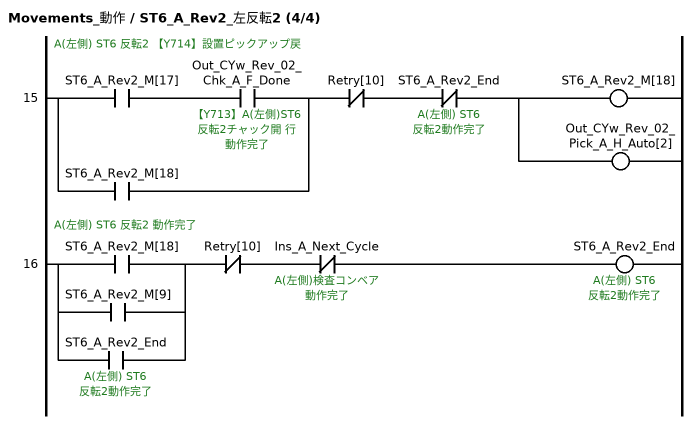
(* [picture p48: Movements_動作 / ST6_A_Rev2_左反転2, rungs 15-16] *)
(* Rung 15: A(左側) ST6 反転2 【Y714】設置ピックアップ戻 *)
_p89 := ((ST6_A_Rev2_M[17] AND Out_CYw_Rev_02_Chk_A_F_Done) OR ST6_A_Rev2_M[18]) AND NOT Retry[10] AND NOT ST6_A_Rev2_End;
ST6_A_Rev2_M[18] := _p89;
Out_CYw_Rev_02_Pick_A_H_Auto[2] := _p89;
(* Rung 16: A(左側) ST6 反転2 動作完了 *)
ST6_A_Rev2_End := (ST6_A_Rev2_M[18] OR ST6_A_Rev2_M[9] OR ST6_A_Rev2_End) AND NOT Retry[10] AND NOT Ins_A_Next_Cycle;

(* Section ST7_A_Dis2_左SF排出: ladder, written here as Structured Text *)

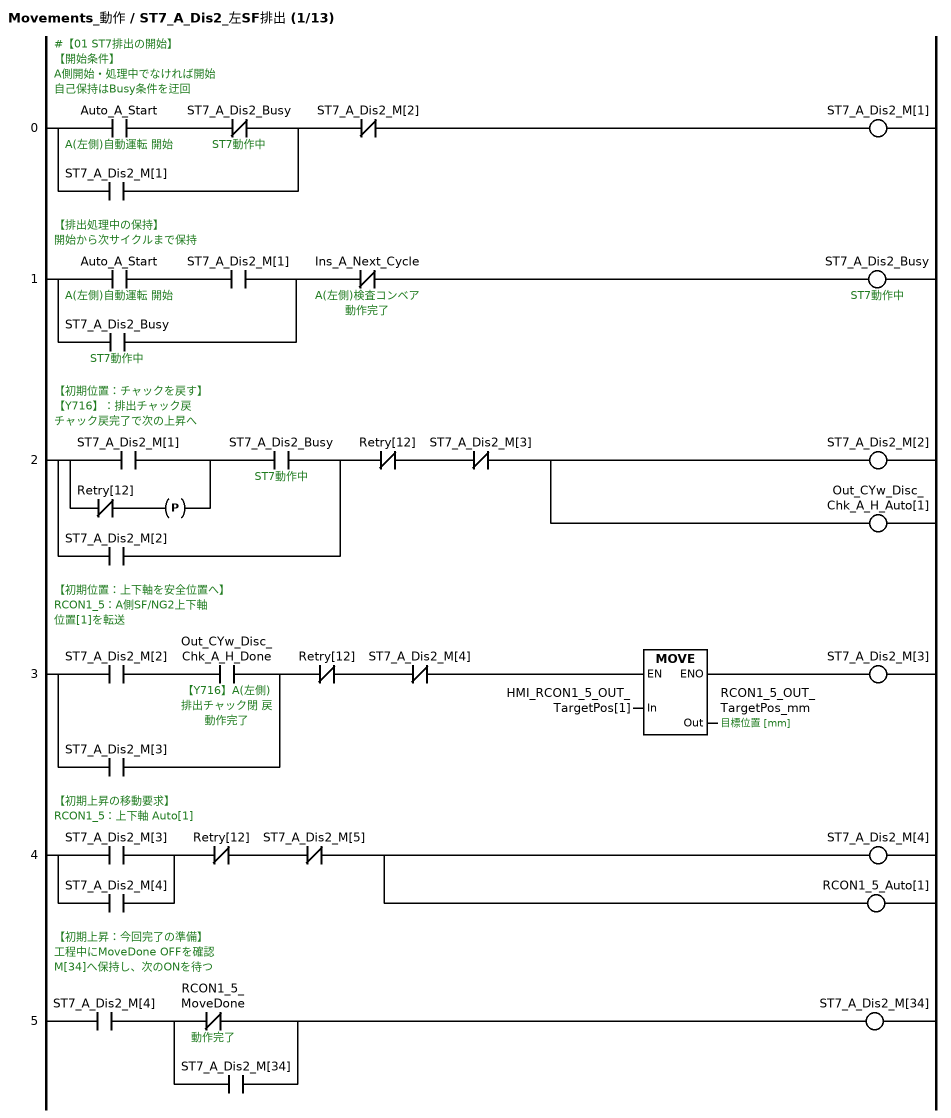
(* Rung 0: #【01 ST7排出の開始】 / 【開始条件】 / A側開始・処理中でなければ開始 / 自己保持はBusy条件を迂回 *)
ST7_A_Dis2_M[1] := ((Auto_A_Start AND NOT ST7_A_Dis2_Busy) OR ST7_A_Dis2_M[1]) AND NOT ST7_A_Dis2_M[2];
(* Rung 1: 【排出処理中の保持】 / 開始から次サイクルまで保持 *)
ST7_A_Dis2_Busy := ((Auto_A_Start AND ST7_A_Dis2_M[1]) OR ST7_A_Dis2_Busy) AND NOT Ins_A_Next_Cycle;
(* Rung 2: 【初期位置：チャックを戻す】 / 【Y716】：排出チャック戻 / チャック戻完了で次の上昇へ *)
_e90(CLK := NOT Retry[12]);
_p91 := (((ST7_A_Dis2_M[1] OR _e90.Q) AND ST7_A_Dis2_Busy) OR ST7_A_Dis2_M[2]) AND NOT Retry[12] AND NOT ST7_A_Dis2_M[3];
ST7_A_Dis2_M[2] := _p91;
Out_CYw_Disc_Chk_A_H_Auto[1] := _p91;
(* Rung 3: 【初期位置：上下軸を安全位置へ】 / RCON1_5：A側SF/NG2上下軸 / 位置[1]を転送 *)
IF ((ST7_A_Dis2_M[2] AND Out_CYw_Disc_Chk_A_H_Done) OR ST7_A_Dis2_M[3]) AND NOT Retry[12] AND NOT ST7_A_Dis2_M[4] THEN
    RCON1_5_OUT_TargetPos_mm := HMI_RCON1_5_OUT_TargetPos[1];
END_IF;
ST7_A_Dis2_M[3] := ((ST7_A_Dis2_M[2] AND Out_CYw_Disc_Chk_A_H_Done) OR ST7_A_Dis2_M[3]) AND NOT Retry[12] AND NOT ST7_A_Dis2_M[4];
(* Rung 4: 【初期上昇の移動要求】 / RCON1_5：上下軸 Auto[1] *)
_p92 := (ST7_A_Dis2_M[3] OR ST7_A_Dis2_M[4]) AND NOT Retry[12] AND NOT ST7_A_Dis2_M[5];
ST7_A_Dis2_M[4] := _p92;
RCON1_5_Auto[1] := _p92;
(* Rung 5: 【初期上昇：今回完了の準備】 / 工程中にMoveDone OFFを確認 / M[34]へ保持し、次のONを待つ *)
ST7_A_Dis2_M[34] := ST7_A_Dis2_M[4] AND (NOT RCON1_5_MoveDone OR ST7_A_Dis2_M[34]);

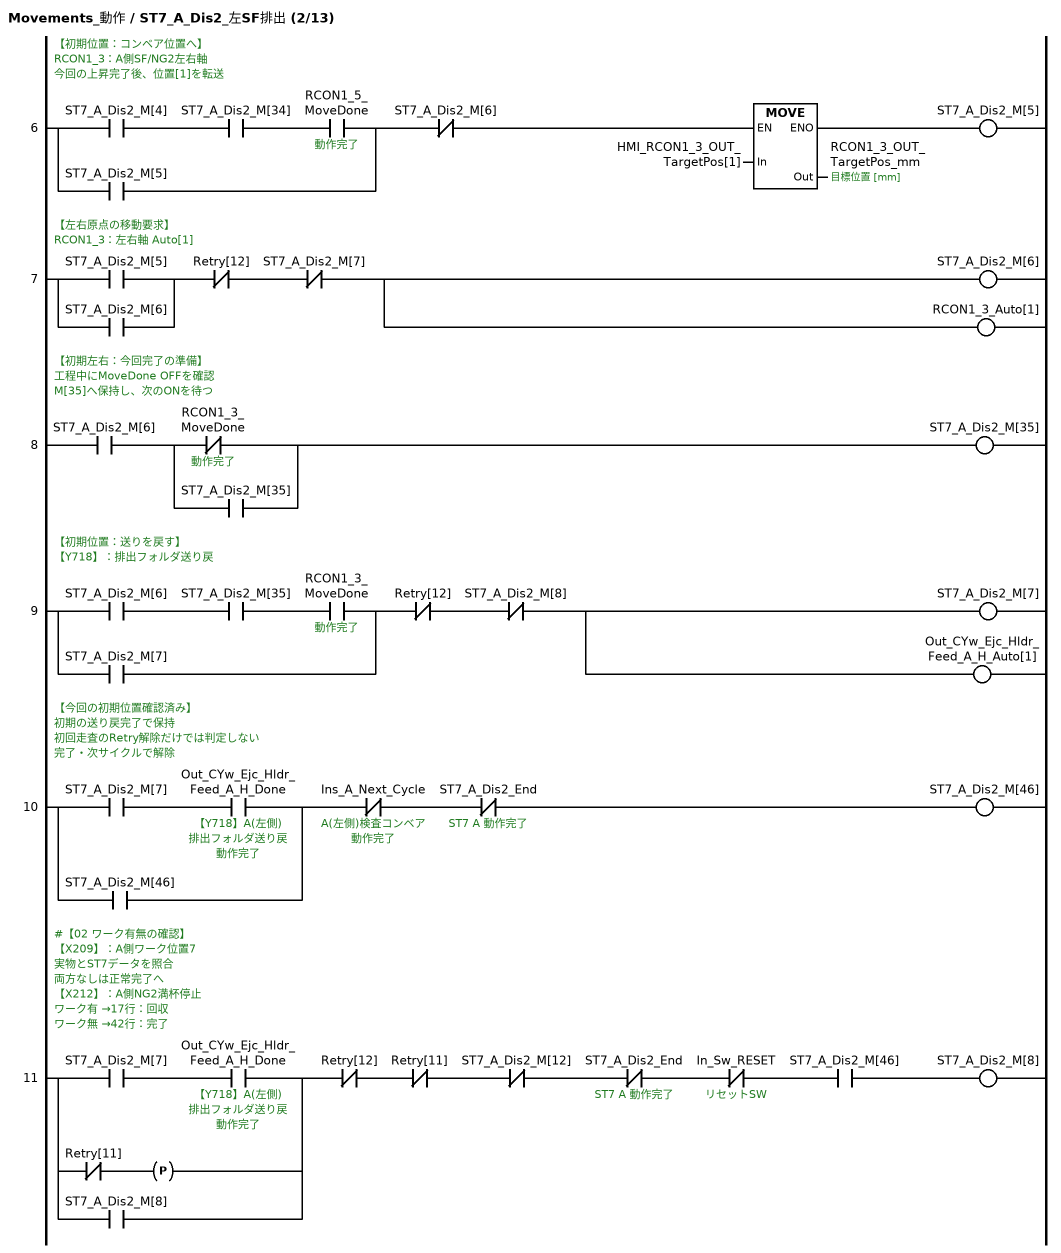
(* Rung 6: 【初期位置：コンベア位置へ】 / RCON1_3：A側SF/NG2左右軸 / 今回の上昇完了後、位置[1]を転送 *)
IF ((ST7_A_Dis2_M[4] AND ST7_A_Dis2_M[34] AND RCON1_5_MoveDone) OR ST7_A_Dis2_M[5]) AND NOT ST7_A_Dis2_M[6] THEN
    RCON1_3_OUT_TargetPos_mm := HMI_RCON1_3_OUT_TargetPos[1];
END_IF;
ST7_A_Dis2_M[5] := ((ST7_A_Dis2_M[4] AND ST7_A_Dis2_M[34] AND RCON1_5_MoveDone) OR ST7_A_Dis2_M[5]) AND NOT ST7_A_Dis2_M[6];
(* Rung 7: 【左右原点の移動要求】 / RCON1_3：左右軸 Auto[1] *)
_p93 := (ST7_A_Dis2_M[5] OR ST7_A_Dis2_M[6]) AND NOT Retry[12] AND NOT ST7_A_Dis2_M[7];
ST7_A_Dis2_M[6] := _p93;
RCON1_3_Auto[1] := _p93;
(* Rung 8: 【初期左右：今回完了の準備】 / 工程中にMoveDone OFFを確認 / M[35]へ保持し、次のONを待つ *)
ST7_A_Dis2_M[35] := ST7_A_Dis2_M[6] AND (NOT RCON1_3_MoveDone OR ST7_A_Dis2_M[35]);
(* Rung 9: 【初期位置：送りを戻す】 / 【Y718】：排出フォルダ送り戻 *)
_p94 := ((ST7_A_Dis2_M[6] AND ST7_A_Dis2_M[35] AND RCON1_3_MoveDone) OR ST7_A_Dis2_M[7]) AND NOT Retry[12] AND NOT ST7_A_Dis2_M[8];
ST7_A_Dis2_M[7] := _p94;
Out_CYw_Ejc_Hldr_Feed_A_H_Auto[1] := _p94;
(* Rung 10: 【今回の初期位置確認済み】 / 初期の送り戻完了で保持 / 初回走査のRetry解除だけでは判定しない / 完了・次サイクルで解除 *)
ST7_A_Dis2_M[46] := ((ST7_A_Dis2_M[7] AND Out_CYw_Ejc_Hldr_Feed_A_H_Done) OR ST7_A_Dis2_M[46]) AND NOT Ins_A_Next_Cycle AND NOT ST7_A_Dis2_End;
(* Rung 11: #【02 ワーク有無の確認】 / 【X209】：A側ワーク位置7 / 実物とST7データを照合 / 両方なしは正常完了へ / 【X212】：A側NG2満杯停止 / ワーク有 →17行：回収 / ワーク無 →42行：完了 *)
_e95(CLK := NOT Retry[11]);
ST7_A_Dis2_M[8] := ((ST7_A_Dis2_M[7] AND Out_CYw_Ejc_Hldr_Feed_A_H_Done) OR _e95.Q OR ST7_A_Dis2_M[8]) AND NOT Retry[12] AND NOT Retry[11] AND NOT ST7_A_Dis2_M[12] AND NOT ST7_A_Dis2_End AND NOT In_Sw_RESET AND ST7_A_Dis2_M[46];

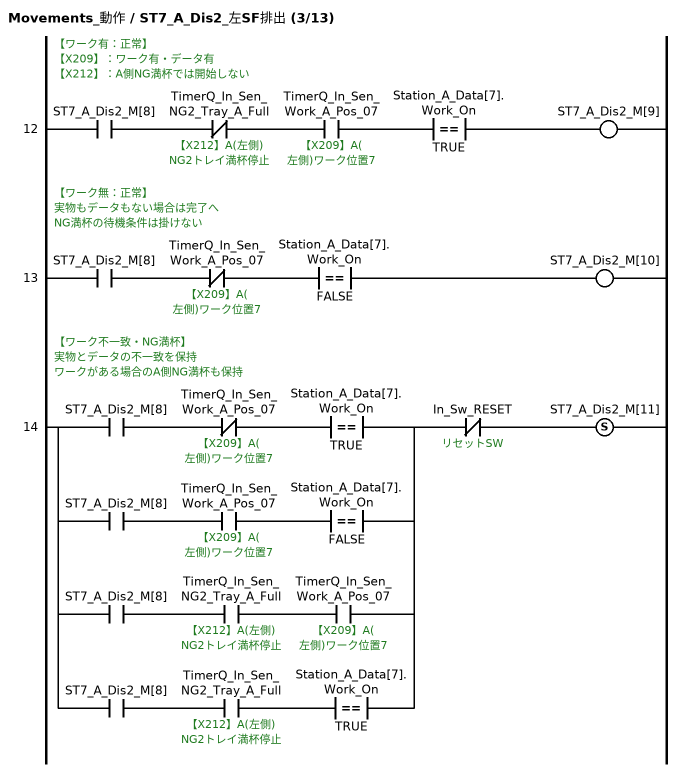
(* Rung 12: 【ワーク有：正常】 / 【X209】：ワーク有・データ有 / 【X212】：A側NG満杯では開始しない *)
ST7_A_Dis2_M[9] := ST7_A_Dis2_M[8] AND NOT TimerQ_In_Sen_NG2_Tray_A_Full AND TimerQ_In_Sen_Work_A_Pos_07 AND (Station_A_Data[7].Work_On = TRUE);
(* Rung 13: 【ワーク無：正常】 / 実物もデータもない場合は完了へ / NG満杯の待機条件は掛けない *)
ST7_A_Dis2_M[10] := ST7_A_Dis2_M[8] AND NOT TimerQ_In_Sen_Work_A_Pos_07 AND (Station_A_Data[7].Work_On = FALSE);
(* Rung 14: 【ワーク不一致・NG満杯】 / 実物とデータの不一致を保持 / ワークがある場合のA側NG満杯も保持 *)
IF ((ST7_A_Dis2_M[8] AND NOT TimerQ_In_Sen_Work_A_Pos_07 AND (Station_A_Data[7].Work_On = TRUE)) OR (ST7_A_Dis2_M[8] AND TimerQ_In_Sen_Work_A_Pos_07 AND (Station_A_Data[7].Work_On = FALSE)) OR (ST7_A_Dis2_M[8] AND TimerQ_In_Sen_NG2_Tray_A_Full AND TimerQ_In_Sen_Work_A_Pos_07) OR (ST7_A_Dis2_M[8] AND TimerQ_In_Sen_NG2_Tray_A_Full AND (Station_A_Data[7].Work_On = TRUE))) AND NOT In_Sw_RESET THEN
    ST7_A_Dis2_M[11] := TRUE;
END_IF;

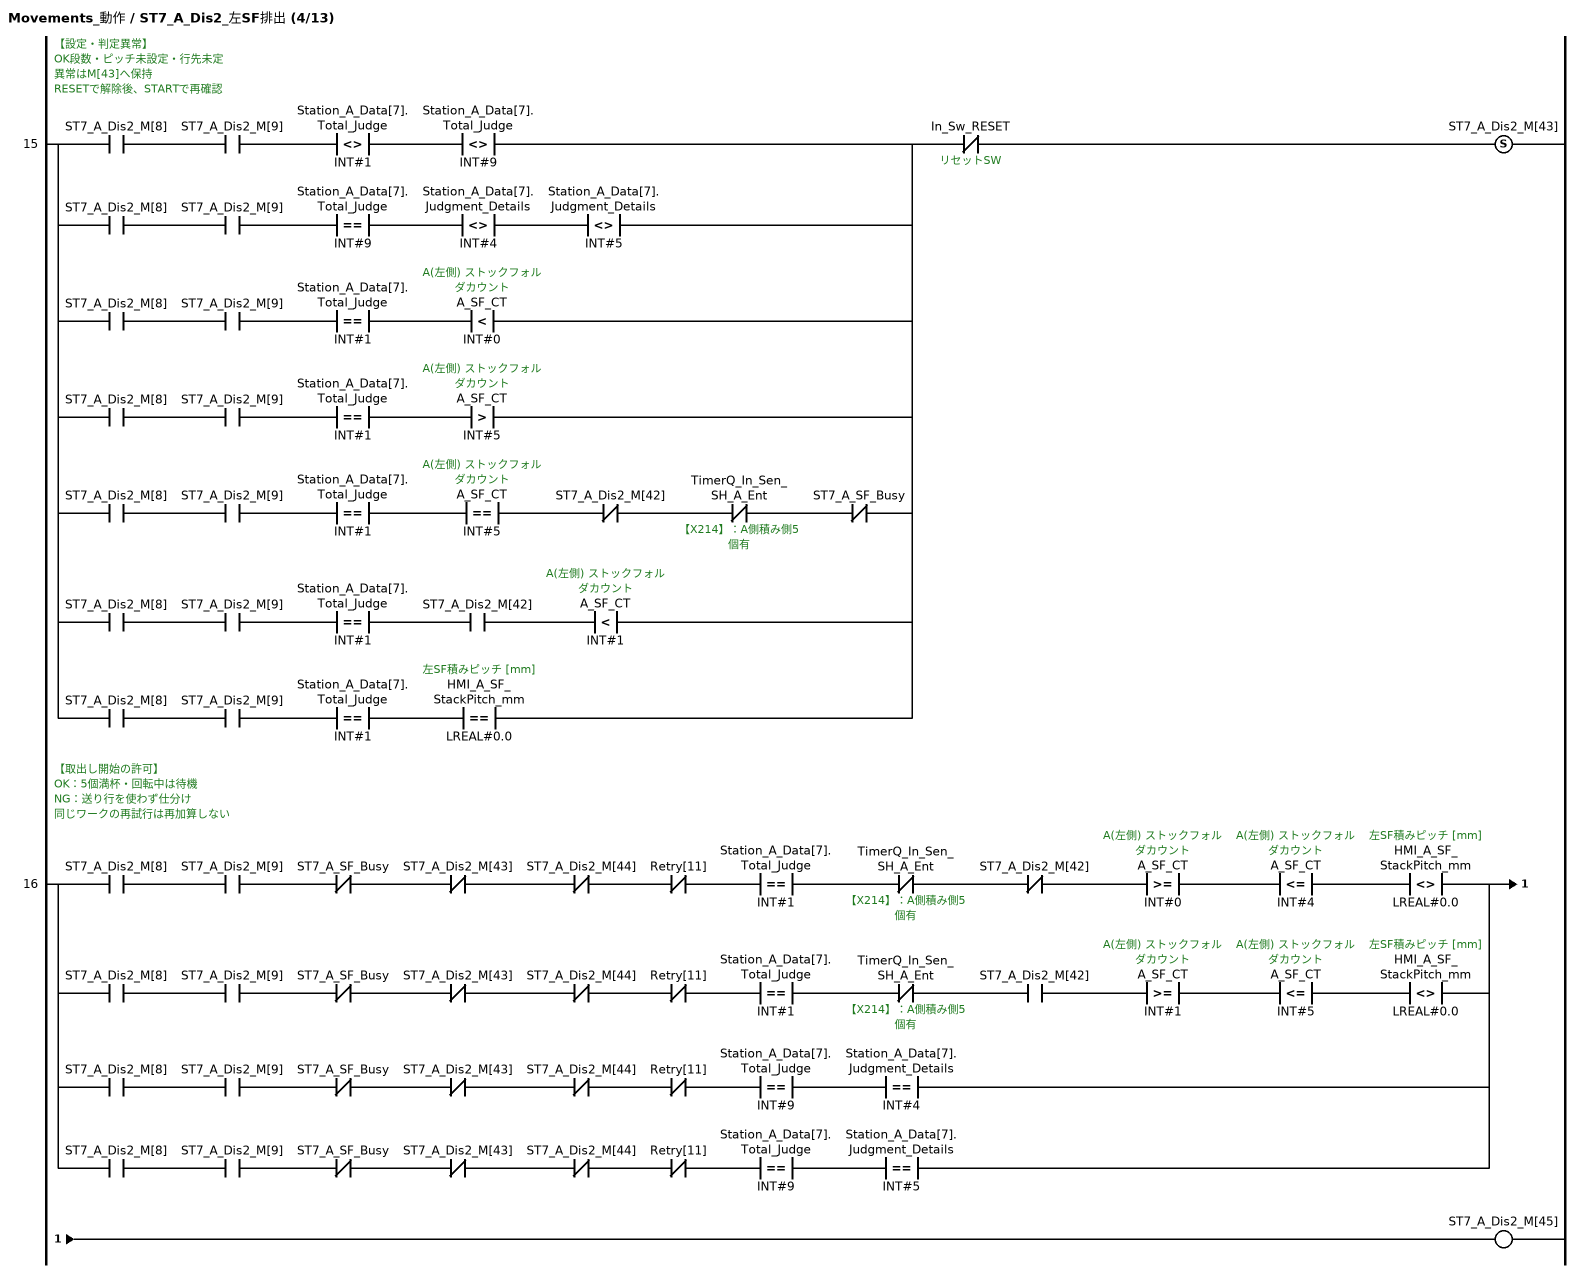
(* Rung 15: 【設定・判定異常】 / OK段数・ピッチ未設定・行先未定 / 異常はM[43]へ保持 / RESETで解除後、STARTで再確認 *)
IF ((ST7_A_Dis2_M[8] AND ST7_A_Dis2_M[9] AND (Station_A_Data[7].Total_Judge <> INT#1) AND (Station_A_Data[7].Total_Judge <> INT#9)) OR (ST7_A_Dis2_M[8] AND ST7_A_Dis2_M[9] AND (Station_A_Data[7].Total_Judge = INT#9) AND (Station_A_Data[7].Judgment_Details <> INT#4) AND (Station_A_Data[7].Judgment_Details <> INT#5)) OR (ST7_A_Dis2_M[8] AND ST7_A_Dis2_M[9] AND (Station_A_Data[7].Total_Judge = INT#1) AND (A_SF_CT < INT#0)) OR (ST7_A_Dis2_M[8] AND ST7_A_Dis2_M[9] AND (Station_A_Data[7].Total_Judge = INT#1) AND (A_SF_CT > INT#5)) OR (ST7_A_Dis2_M[8] AND ST7_A_Dis2_M[9] AND (Station_A_Data[7].Total_Judge = INT#1) AND (A_SF_CT = INT#5) AND NOT ST7_A_Dis2_M[42] AND NOT TimerQ_In_Sen_SH_A_Ent AND NOT ST7_A_SF_Busy) OR (ST7_A_Dis2_M[8] AND ST7_A_Dis2_M[9] AND (Station_A_Data[7].Total_Judge = INT#1) AND ST7_A_Dis2_M[42] AND (A_SF_CT < INT#1)) OR (ST7_A_Dis2_M[8] AND ST7_A_Dis2_M[9] AND (Station_A_Data[7].Total_Judge = INT#1) AND (HMI_A_SF_StackPitch_mm = LREAL#0.0))) AND NOT In_Sw_RESET THEN
    ST7_A_Dis2_M[43] := TRUE;
END_IF;
(* Rung 16: 【取出し開始の許可】 / OK：5個満杯・回転中は待機 / NG：送り行を使わず仕分け / 同じワークの再試行は再加算しない *)
ST7_A_Dis2_M[45] := (ST7_A_Dis2_M[8] AND ST7_A_Dis2_M[9] AND NOT ST7_A_SF_Busy AND NOT ST7_A_Dis2_M[43] AND NOT ST7_A_Dis2_M[44] AND NOT Retry[11] AND (Station_A_Data[7].Total_Judge = INT#1) AND NOT TimerQ_In_Sen_SH_A_Ent AND NOT ST7_A_Dis2_M[42] AND (A_SF_CT >= INT#0) AND (A_SF_CT <= INT#4) AND (HMI_A_SF_StackPitch_mm <> LREAL#0.0)) OR (ST7_A_Dis2_M[8] AND ST7_A_Dis2_M[9] AND NOT ST7_A_SF_Busy AND NOT ST7_A_Dis2_M[43] AND NOT ST7_A_Dis2_M[44] AND NOT Retry[11] AND (Station_A_Data[7].Total_Judge = INT#1) AND NOT TimerQ_In_Sen_SH_A_Ent AND ST7_A_Dis2_M[42] AND (A_SF_CT >= INT#1) AND (A_SF_CT <= INT#5) AND (HMI_A_SF_StackPitch_mm <> LREAL#0.0)) OR (ST7_A_Dis2_M[8] AND ST7_A_Dis2_M[9] AND NOT ST7_A_SF_Busy AND NOT ST7_A_Dis2_M[43] AND NOT ST7_A_Dis2_M[44] AND NOT Retry[11] AND (Station_A_Data[7].Total_Judge = INT#9) AND (Station_A_Data[7].Judgment_Details = INT#4)) OR (ST7_A_Dis2_M[8] AND ST7_A_Dis2_M[9] AND NOT ST7_A_SF_Busy AND NOT ST7_A_Dis2_M[43] AND NOT ST7_A_Dis2_M[44] AND NOT Retry[11] AND (Station_A_Data[7].Total_Judge = INT#9) AND (Station_A_Data[7].Judgment_Details = INT#5));

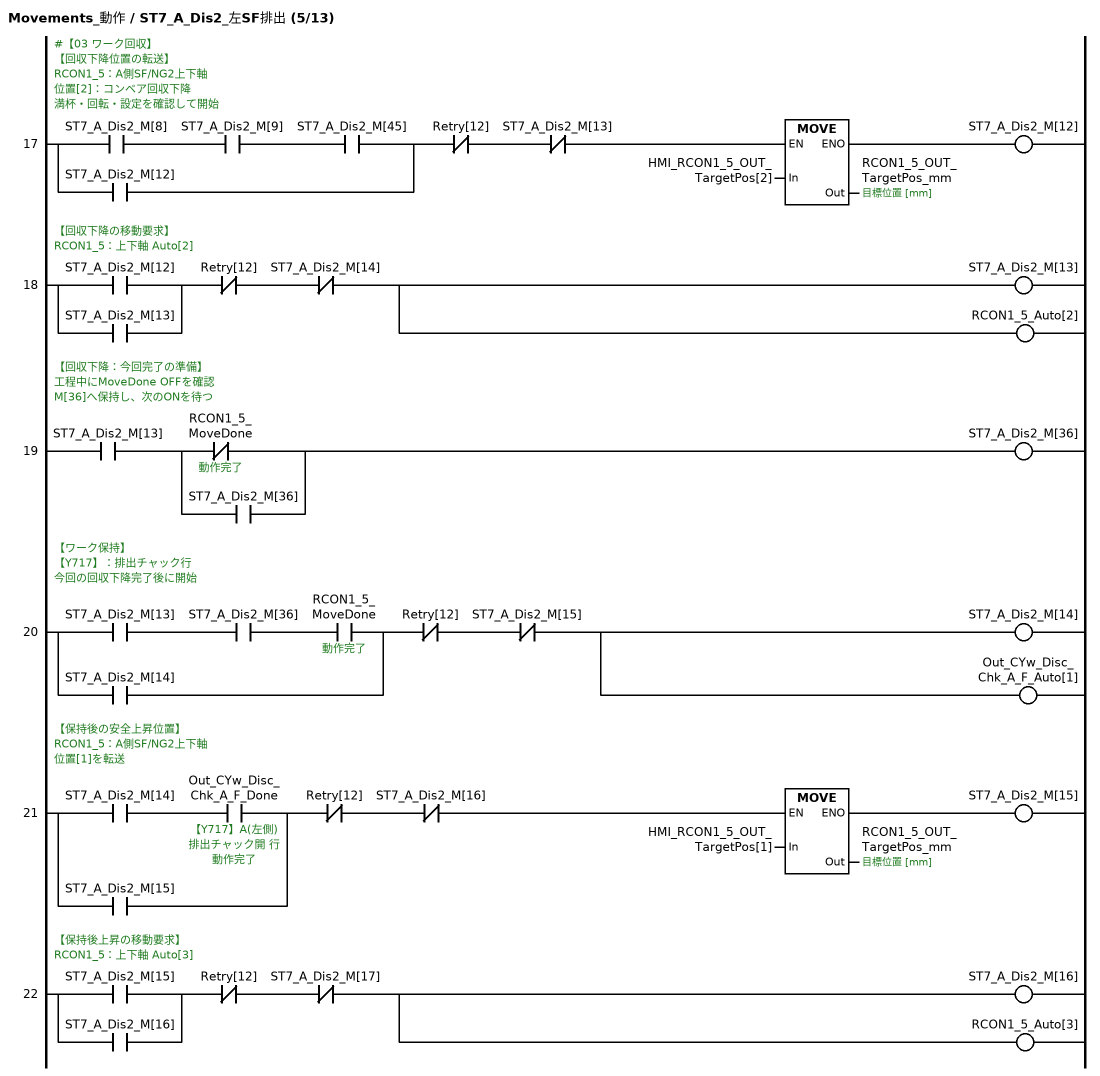
(* Rung 17: #【03 ワーク回収】 / 【回収下降位置の転送】 / RCON1_5：A側SF/NG2上下軸 / 位置[2]：コンベア回収下降 / 満杯・回転・設定を確認して開始 *)
IF ((ST7_A_Dis2_M[8] AND ST7_A_Dis2_M[9] AND ST7_A_Dis2_M[45]) OR ST7_A_Dis2_M[12]) AND NOT Retry[12] AND NOT ST7_A_Dis2_M[13] THEN
    RCON1_5_OUT_TargetPos_mm := HMI_RCON1_5_OUT_TargetPos[2];
END_IF;
ST7_A_Dis2_M[12] := ((ST7_A_Dis2_M[8] AND ST7_A_Dis2_M[9] AND ST7_A_Dis2_M[45]) OR ST7_A_Dis2_M[12]) AND NOT Retry[12] AND NOT ST7_A_Dis2_M[13];
(* Rung 18: 【回収下降の移動要求】 / RCON1_5：上下軸 Auto[2] *)
_p96 := (ST7_A_Dis2_M[12] OR ST7_A_Dis2_M[13]) AND NOT Retry[12] AND NOT ST7_A_Dis2_M[14];
ST7_A_Dis2_M[13] := _p96;
RCON1_5_Auto[2] := _p96;
(* Rung 19: 【回収下降：今回完了の準備】 / 工程中にMoveDone OFFを確認 / M[36]へ保持し、次のONを待つ *)
ST7_A_Dis2_M[36] := ST7_A_Dis2_M[13] AND (NOT RCON1_5_MoveDone OR ST7_A_Dis2_M[36]);
(* Rung 20: 【ワーク保持】 / 【Y717】：排出チャック行 / 今回の回収下降完了後に開始 *)
_p97 := ((ST7_A_Dis2_M[13] AND ST7_A_Dis2_M[36] AND RCON1_5_MoveDone) OR ST7_A_Dis2_M[14]) AND NOT Retry[12] AND NOT ST7_A_Dis2_M[15];
ST7_A_Dis2_M[14] := _p97;
Out_CYw_Disc_Chk_A_F_Auto[1] := _p97;
(* Rung 21: 【保持後の安全上昇位置】 / RCON1_5：A側SF/NG2上下軸 / 位置[1]を転送 *)
IF ((ST7_A_Dis2_M[14] AND Out_CYw_Disc_Chk_A_F_Done) OR ST7_A_Dis2_M[15]) AND NOT Retry[12] AND NOT ST7_A_Dis2_M[16] THEN
    RCON1_5_OUT_TargetPos_mm := HMI_RCON1_5_OUT_TargetPos[1];
END_IF;
ST7_A_Dis2_M[15] := ((ST7_A_Dis2_M[14] AND Out_CYw_Disc_Chk_A_F_Done) OR ST7_A_Dis2_M[15]) AND NOT Retry[12] AND NOT ST7_A_Dis2_M[16];
(* Rung 22: 【保持後上昇の移動要求】 / RCON1_5：上下軸 Auto[3] *)
_p98 := (ST7_A_Dis2_M[15] OR ST7_A_Dis2_M[16]) AND NOT Retry[12] AND NOT ST7_A_Dis2_M[17];
ST7_A_Dis2_M[16] := _p98;
RCON1_5_Auto[3] := _p98;

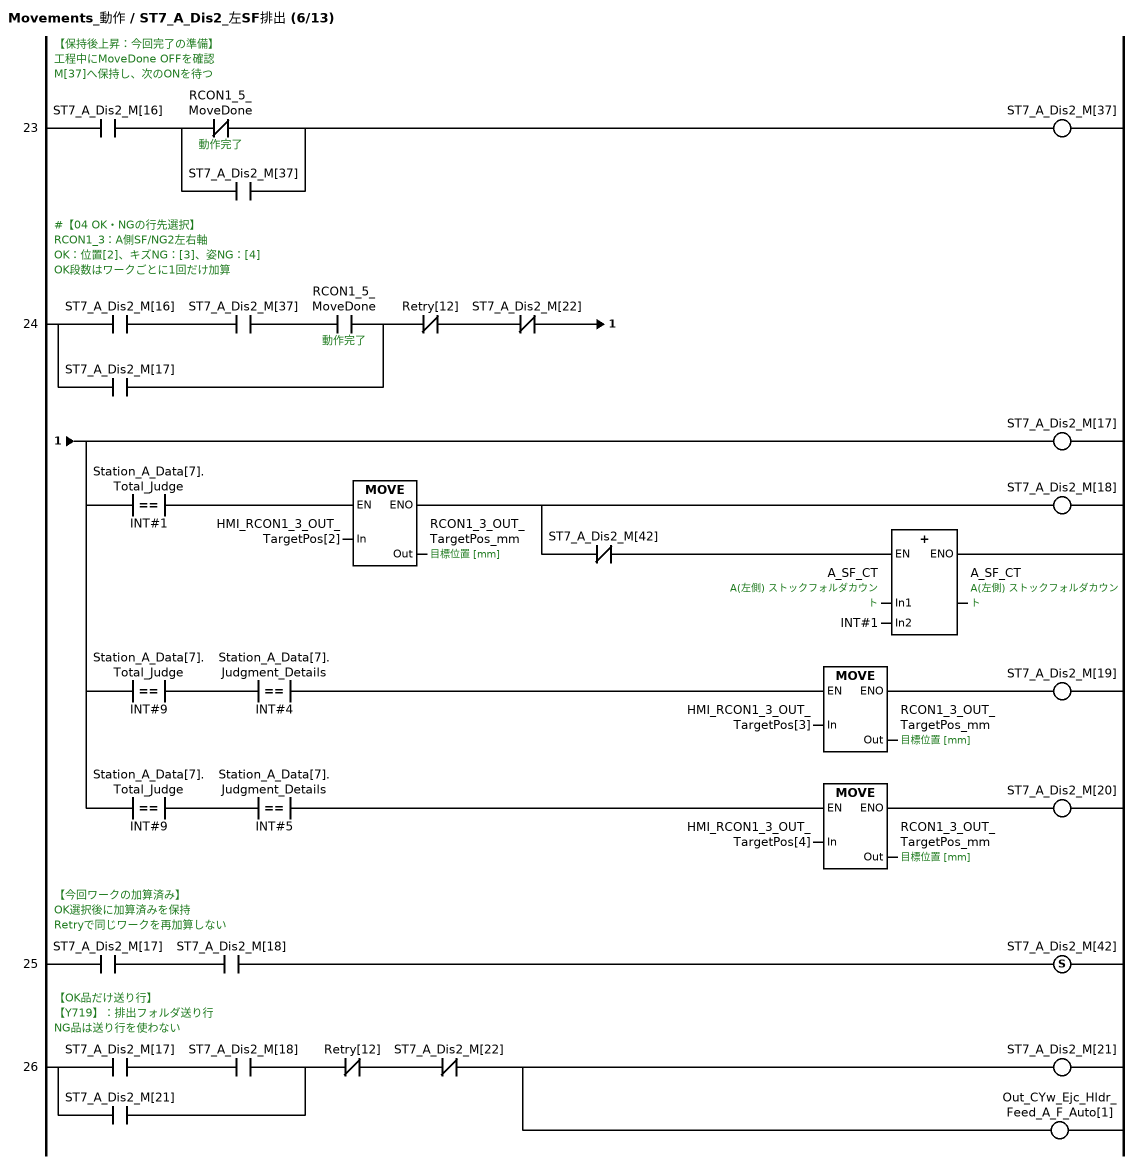
(* Rung 23: 【保持後上昇：今回完了の準備】 / 工程中にMoveDone OFFを確認 / M[37]へ保持し、次のONを待つ *)
ST7_A_Dis2_M[37] := ST7_A_Dis2_M[16] AND (NOT RCON1_5_MoveDone OR ST7_A_Dis2_M[37]);
(* Rung 24: #【04 OK・NGの行先選択】 / RCON1_3：A側SF/NG2左右軸 / OK：位置[2]、キズNG：[3]、姿NG：[4] / OK段数はワークごとに1回だけ加算 *)
_p99 := ((ST7_A_Dis2_M[16] AND ST7_A_Dis2_M[37] AND RCON1_5_MoveDone) OR ST7_A_Dis2_M[17]) AND NOT Retry[12] AND NOT ST7_A_Dis2_M[22];
ST7_A_Dis2_M[17] := _p99;
IF _p99 AND (Station_A_Data[7].Total_Judge = INT#1) THEN
    RCON1_3_OUT_TargetPos_mm := HMI_RCON1_3_OUT_TargetPos[2];
END_IF;
ST7_A_Dis2_M[18] := _p99 AND (Station_A_Data[7].Total_Judge = INT#1);
IF _p99 AND (Station_A_Data[7].Total_Judge = INT#1) AND NOT ST7_A_Dis2_M[42] THEN
    A_SF_CT := A_SF_CT + INT#1;
END_IF;
IF _p99 AND (Station_A_Data[7].Total_Judge = INT#9) AND (Station_A_Data[7].Judgment_Details = INT#4) THEN
    RCON1_3_OUT_TargetPos_mm := HMI_RCON1_3_OUT_TargetPos[3];
END_IF;
ST7_A_Dis2_M[19] := _p99 AND (Station_A_Data[7].Total_Judge = INT#9) AND (Station_A_Data[7].Judgment_Details = INT#4);
IF _p99 AND (Station_A_Data[7].Total_Judge = INT#9) AND (Station_A_Data[7].Judgment_Details = INT#5) THEN
    RCON1_3_OUT_TargetPos_mm := HMI_RCON1_3_OUT_TargetPos[4];
END_IF;
ST7_A_Dis2_M[20] := _p99 AND (Station_A_Data[7].Total_Judge = INT#9) AND (Station_A_Data[7].Judgment_Details = INT#5);
(* Rung 25: 【今回ワークの加算済み】 / OK選択後に加算済みを保持 / Retryで同じワークを再加算しない *)
IF ST7_A_Dis2_M[17] AND ST7_A_Dis2_M[18] THEN ST7_A_Dis2_M[42] := TRUE; END_IF;
(* Rung 26: 【OK品だけ送り行】 / 【Y719】：排出フォルダ送り行 / NG品は送り行を使わない *)
_p100 := ((ST7_A_Dis2_M[17] AND ST7_A_Dis2_M[18]) OR ST7_A_Dis2_M[21]) AND NOT Retry[12] AND NOT ST7_A_Dis2_M[22];
ST7_A_Dis2_M[21] := _p100;
Out_CYw_Ejc_Hldr_Feed_A_F_Auto[1] := _p100;

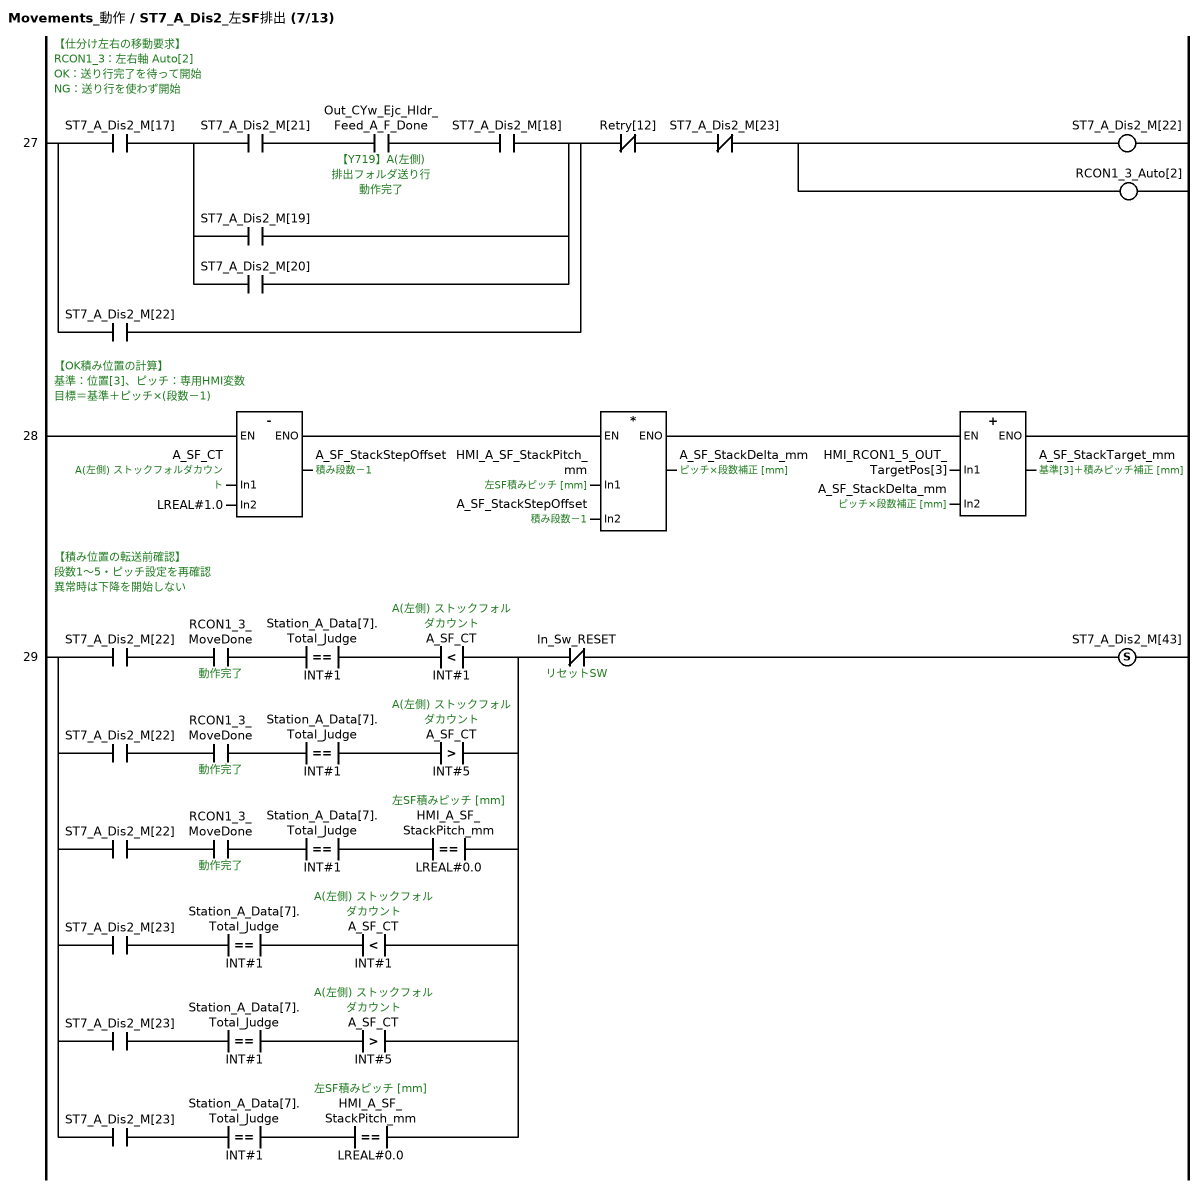
(* Rung 27: 【仕分け左右の移動要求】 / RCON1_3：左右軸 Auto[2] / OK：送り行完了を待って開始 / NG：送り行を使わず開始 *)
_p101 := ((ST7_A_Dis2_M[17] AND ((ST7_A_Dis2_M[21] AND Out_CYw_Ejc_Hldr_Feed_A_F_Done AND ST7_A_Dis2_M[18]) OR ST7_A_Dis2_M[19] OR ST7_A_Dis2_M[20])) OR ST7_A_Dis2_M[22]) AND NOT Retry[12] AND NOT ST7_A_Dis2_M[23];
ST7_A_Dis2_M[22] := _p101;
RCON1_3_Auto[2] := _p101;
(* Rung 28: 【OK積み位置の計算】 / 基準：位置[3]、ピッチ：専用HMI変数 / 目標＝基準＋ピッチ×(段数－1) *)
A_SF_StackStepOffset := A_SF_CT - LREAL#1.0;
A_SF_StackDelta_mm := HMI_A_SF_StackPitch_mm * A_SF_StackStepOffset;
A_SF_StackTarget_mm := HMI_RCON1_5_OUT_TargetPos[3] + A_SF_StackDelta_mm;
(* Rung 29: 【積み位置の転送前確認】 / 段数1～5・ピッチ設定を再確認 / 異常時は下降を開始しない *)
IF ((ST7_A_Dis2_M[22] AND RCON1_3_MoveDone AND (Station_A_Data[7].Total_Judge = INT#1) AND (A_SF_CT < INT#1)) OR (ST7_A_Dis2_M[22] AND RCON1_3_MoveDone AND (Station_A_Data[7].Total_Judge = INT#1) AND (A_SF_CT > INT#5)) OR (ST7_A_Dis2_M[22] AND RCON1_3_MoveDone AND (Station_A_Data[7].Total_Judge = INT#1) AND (HMI_A_SF_StackPitch_mm = LREAL#0.0)) OR (ST7_A_Dis2_M[23] AND (Station_A_Data[7].Total_Judge = INT#1) AND (A_SF_CT < INT#1)) OR (ST7_A_Dis2_M[23] AND (Station_A_Data[7].Total_Judge = INT#1) AND (A_SF_CT > INT#5)) OR (ST7_A_Dis2_M[23] AND (Station_A_Data[7].Total_Judge = INT#1) AND (HMI_A_SF_StackPitch_mm = LREAL#0.0))) AND NOT In_Sw_RESET THEN
    ST7_A_Dis2_M[43] := TRUE;
END_IF;

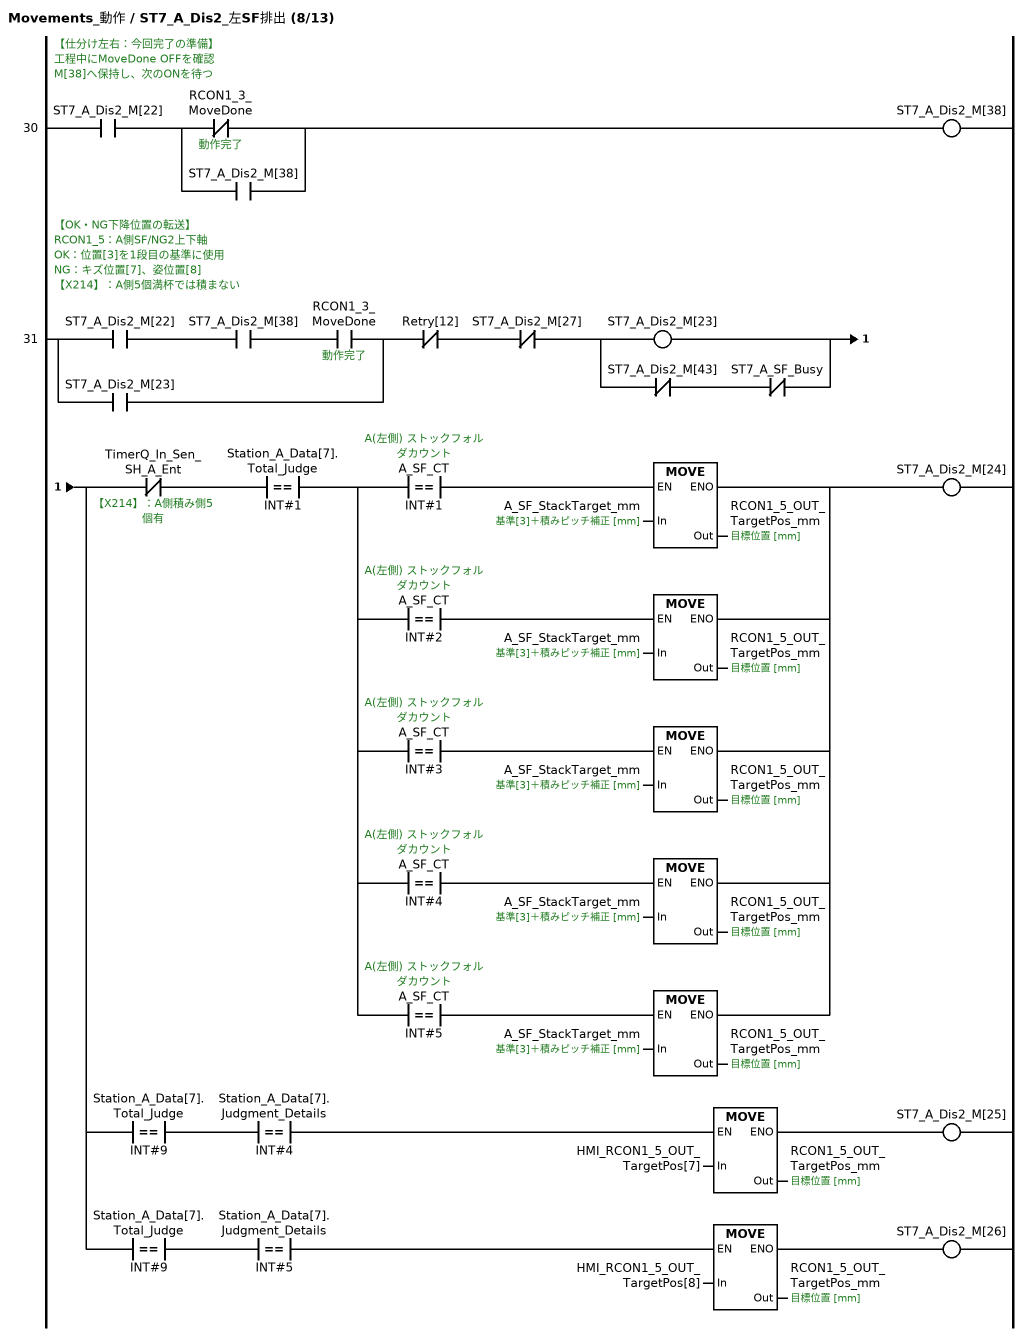
(* Rung 30: 【仕分け左右：今回完了の準備】 / 工程中にMoveDone OFFを確認 / M[38]へ保持し、次のONを待つ *)
ST7_A_Dis2_M[38] := ST7_A_Dis2_M[22] AND (NOT RCON1_3_MoveDone OR ST7_A_Dis2_M[38]);
(* Rung 31: 【OK・NG下降位置の転送】 / RCON1_5：A側SF/NG2上下軸 / OK：位置[3]を1段目の基準に使用 / NG：キズ位置[7]、姿位置[8] / 【X214】：A側5個満杯では積まない *)
_p102 := ((ST7_A_Dis2_M[22] AND ST7_A_Dis2_M[38] AND RCON1_3_MoveDone) OR ST7_A_Dis2_M[23]) AND NOT Retry[12] AND NOT ST7_A_Dis2_M[27];
ST7_A_Dis2_M[23] := _p102;
_p103 := _p102 OR (_p102 AND NOT ST7_A_Dis2_M[43] AND NOT ST7_A_SF_Busy);
_p104 := _p103 AND NOT TimerQ_In_Sen_SH_A_Ent AND (Station_A_Data[7].Total_Judge = INT#1);
IF _p104 AND (A_SF_CT = INT#1) THEN RCON1_5_OUT_TargetPos_mm := A_SF_StackTarget_mm; END_IF;
IF _p104 AND (A_SF_CT = INT#2) THEN RCON1_5_OUT_TargetPos_mm := A_SF_StackTarget_mm; END_IF;
IF _p104 AND (A_SF_CT = INT#3) THEN RCON1_5_OUT_TargetPos_mm := A_SF_StackTarget_mm; END_IF;
IF _p104 AND (A_SF_CT = INT#4) THEN RCON1_5_OUT_TargetPos_mm := A_SF_StackTarget_mm; END_IF;
IF _p104 AND (A_SF_CT = INT#5) THEN RCON1_5_OUT_TargetPos_mm := A_SF_StackTarget_mm; END_IF;
ST7_A_Dis2_M[24] := _p104 AND ((A_SF_CT = INT#1) OR (A_SF_CT = INT#2) OR (A_SF_CT = INT#3) OR (A_SF_CT = INT#4) OR (A_SF_CT = INT#5));
IF _p103 AND (Station_A_Data[7].Total_Judge = INT#9) AND (Station_A_Data[7].Judgment_Details = INT#4) THEN
    RCON1_5_OUT_TargetPos_mm := HMI_RCON1_5_OUT_TargetPos[7];
END_IF;
ST7_A_Dis2_M[25] := _p103 AND (Station_A_Data[7].Total_Judge = INT#9) AND (Station_A_Data[7].Judgment_Details = INT#4);
IF _p103 AND (Station_A_Data[7].Total_Judge = INT#9) AND (Station_A_Data[7].Judgment_Details = INT#5) THEN
    RCON1_5_OUT_TargetPos_mm := HMI_RCON1_5_OUT_TargetPos[8];
END_IF;
ST7_A_Dis2_M[26] := _p103 AND (Station_A_Data[7].Total_Judge = INT#9) AND (Station_A_Data[7].Judgment_Details = INT#5);

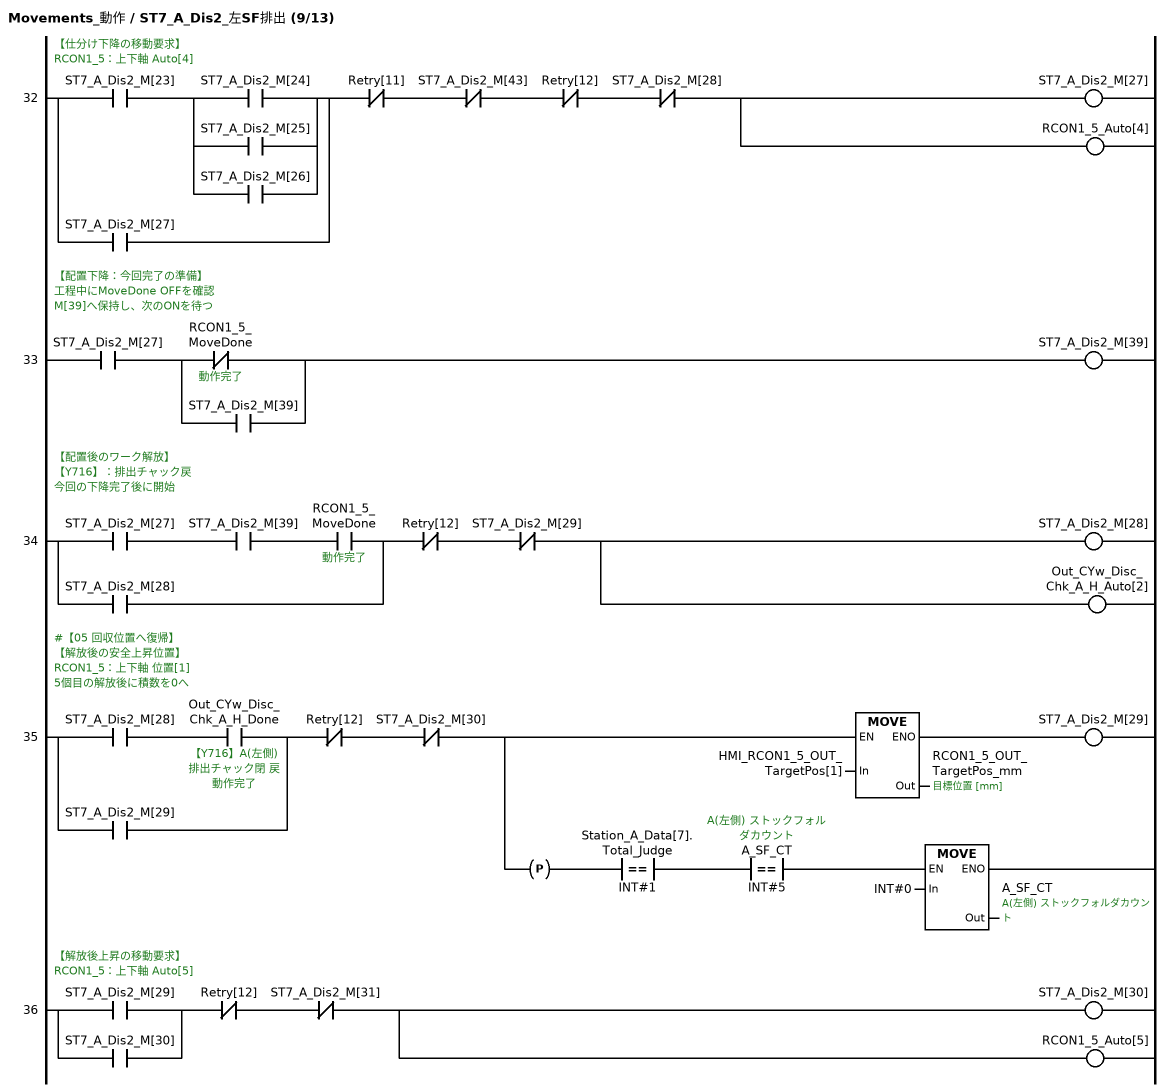
(* Rung 32: 【仕分け下降の移動要求】 / RCON1_5：上下軸 Auto[4] *)
_p105 := ((ST7_A_Dis2_M[23] AND (ST7_A_Dis2_M[24] OR ST7_A_Dis2_M[25] OR ST7_A_Dis2_M[26])) OR ST7_A_Dis2_M[27]) AND NOT Retry[11] AND NOT ST7_A_Dis2_M[43] AND NOT Retry[12] AND NOT ST7_A_Dis2_M[28];
ST7_A_Dis2_M[27] := _p105;
RCON1_5_Auto[4] := _p105;
(* Rung 33: 【配置下降：今回完了の準備】 / 工程中にMoveDone OFFを確認 / M[39]へ保持し、次のONを待つ *)
ST7_A_Dis2_M[39] := ST7_A_Dis2_M[27] AND (NOT RCON1_5_MoveDone OR ST7_A_Dis2_M[39]);
(* Rung 34: 【配置後のワーク解放】 / 【Y716】：排出チャック戻 / 今回の下降完了後に開始 *)
_p106 := ((ST7_A_Dis2_M[27] AND ST7_A_Dis2_M[39] AND RCON1_5_MoveDone) OR ST7_A_Dis2_M[28]) AND NOT Retry[12] AND NOT ST7_A_Dis2_M[29];
ST7_A_Dis2_M[28] := _p106;
Out_CYw_Disc_Chk_A_H_Auto[2] := _p106;
(* Rung 35: #【05 回収位置へ復帰】 / 【解放後の安全上昇位置】 / RCON1_5：上下軸 位置[1] / 5個目の解放後に積数を0へ *)
_p107 := ((ST7_A_Dis2_M[28] AND Out_CYw_Disc_Chk_A_H_Done) OR ST7_A_Dis2_M[29]) AND NOT Retry[12] AND NOT ST7_A_Dis2_M[30];
IF _p107 THEN RCON1_5_OUT_TargetPos_mm := HMI_RCON1_5_OUT_TargetPos[1]; END_IF;
ST7_A_Dis2_M[29] := _p107;
_e108(CLK := _p107);
IF _e108.Q AND (Station_A_Data[7].Total_Judge = INT#1) AND (A_SF_CT = INT#5) THEN
    A_SF_CT := INT#0;
END_IF;
(* Rung 36: 【解放後上昇の移動要求】 / RCON1_5：上下軸 Auto[5] *)
_p109 := (ST7_A_Dis2_M[29] OR ST7_A_Dis2_M[30]) AND NOT Retry[12] AND NOT ST7_A_Dis2_M[31];
ST7_A_Dis2_M[30] := _p109;
RCON1_5_Auto[5] := _p109;

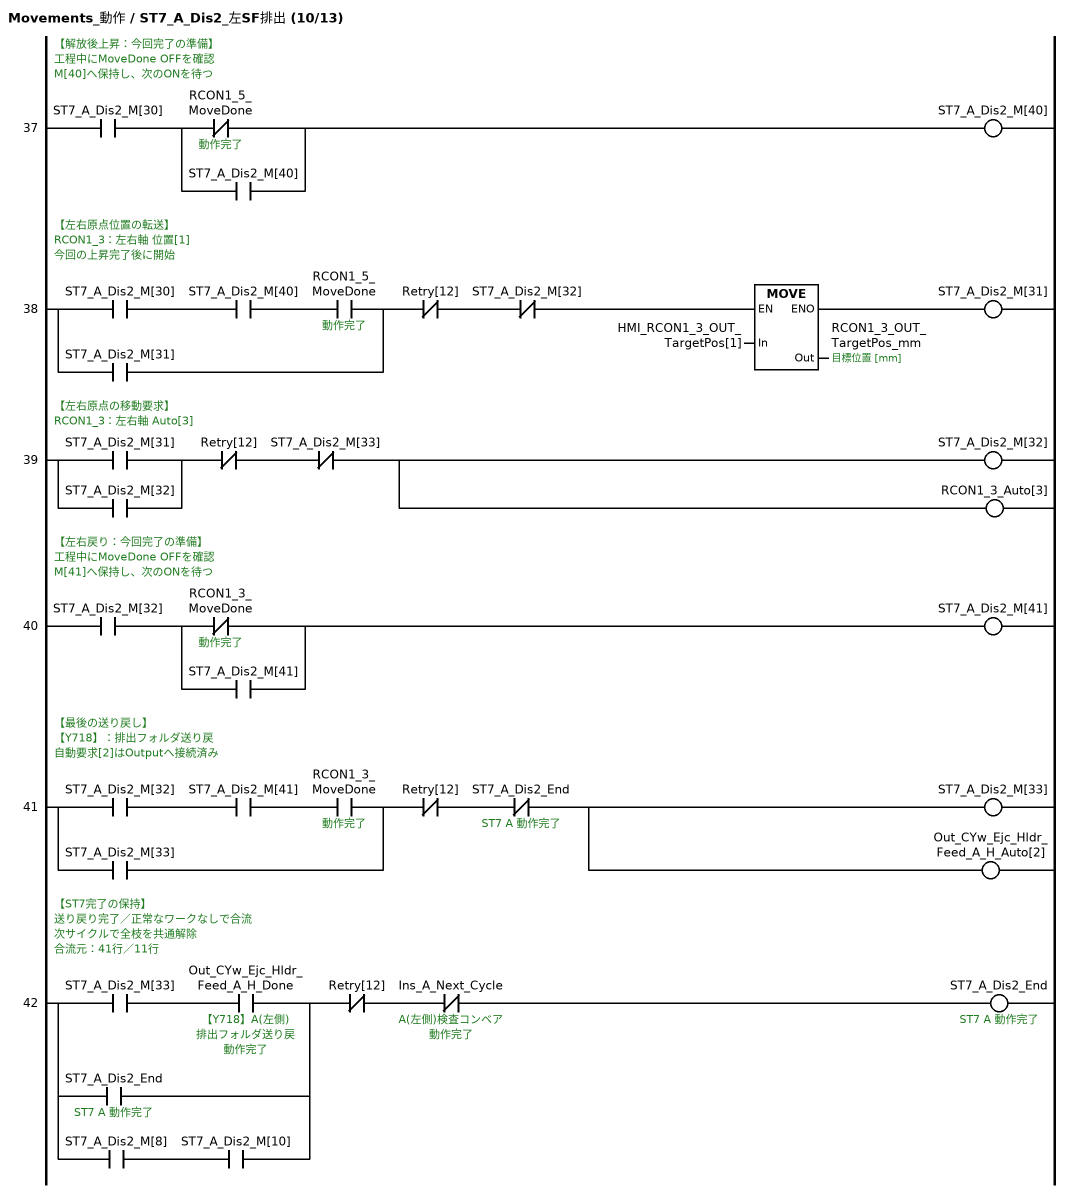
(* Rung 37: 【解放後上昇：今回完了の準備】 / 工程中にMoveDone OFFを確認 / M[40]へ保持し、次のONを待つ *)
ST7_A_Dis2_M[40] := ST7_A_Dis2_M[30] AND (NOT RCON1_5_MoveDone OR ST7_A_Dis2_M[40]);
(* Rung 38: 【左右原点位置の転送】 / RCON1_3：左右軸 位置[1] / 今回の上昇完了後に開始 *)
IF ((ST7_A_Dis2_M[30] AND ST7_A_Dis2_M[40] AND RCON1_5_MoveDone) OR ST7_A_Dis2_M[31]) AND NOT Retry[12] AND NOT ST7_A_Dis2_M[32] THEN
    RCON1_3_OUT_TargetPos_mm := HMI_RCON1_3_OUT_TargetPos[1];
END_IF;
ST7_A_Dis2_M[31] := ((ST7_A_Dis2_M[30] AND ST7_A_Dis2_M[40] AND RCON1_5_MoveDone) OR ST7_A_Dis2_M[31]) AND NOT Retry[12] AND NOT ST7_A_Dis2_M[32];
(* Rung 39: 【左右原点の移動要求】 / RCON1_3：左右軸 Auto[3] *)
_p110 := (ST7_A_Dis2_M[31] OR ST7_A_Dis2_M[32]) AND NOT Retry[12] AND NOT ST7_A_Dis2_M[33];
ST7_A_Dis2_M[32] := _p110;
RCON1_3_Auto[3] := _p110;
(* Rung 40: 【左右戻り：今回完了の準備】 / 工程中にMoveDone OFFを確認 / M[41]へ保持し、次のONを待つ *)
ST7_A_Dis2_M[41] := ST7_A_Dis2_M[32] AND (NOT RCON1_3_MoveDone OR ST7_A_Dis2_M[41]);
(* Rung 41: 【最後の送り戻し】 / 【Y718】：排出フォルダ送り戻 / 自動要求[2]はOutputへ接続済み *)
_p111 := ((ST7_A_Dis2_M[32] AND ST7_A_Dis2_M[41] AND RCON1_3_MoveDone) OR ST7_A_Dis2_M[33]) AND NOT Retry[12] AND NOT ST7_A_Dis2_End;
ST7_A_Dis2_M[33] := _p111;
Out_CYw_Ejc_Hldr_Feed_A_H_Auto[2] := _p111;
(* Rung 42: 【ST7完了の保持】 / 送り戻り完了／正常なワークなしで合流 / 次サイクルで全枝を共通解除 / 合流元：41行／11行 *)
ST7_A_Dis2_End := ((ST7_A_Dis2_M[33] AND Out_CYw_Ejc_Hldr_Feed_A_H_Done) OR ST7_A_Dis2_End OR (ST7_A_Dis2_M[8] AND ST7_A_Dis2_M[10])) AND NOT Retry[12] AND NOT Ins_A_Next_Cycle;

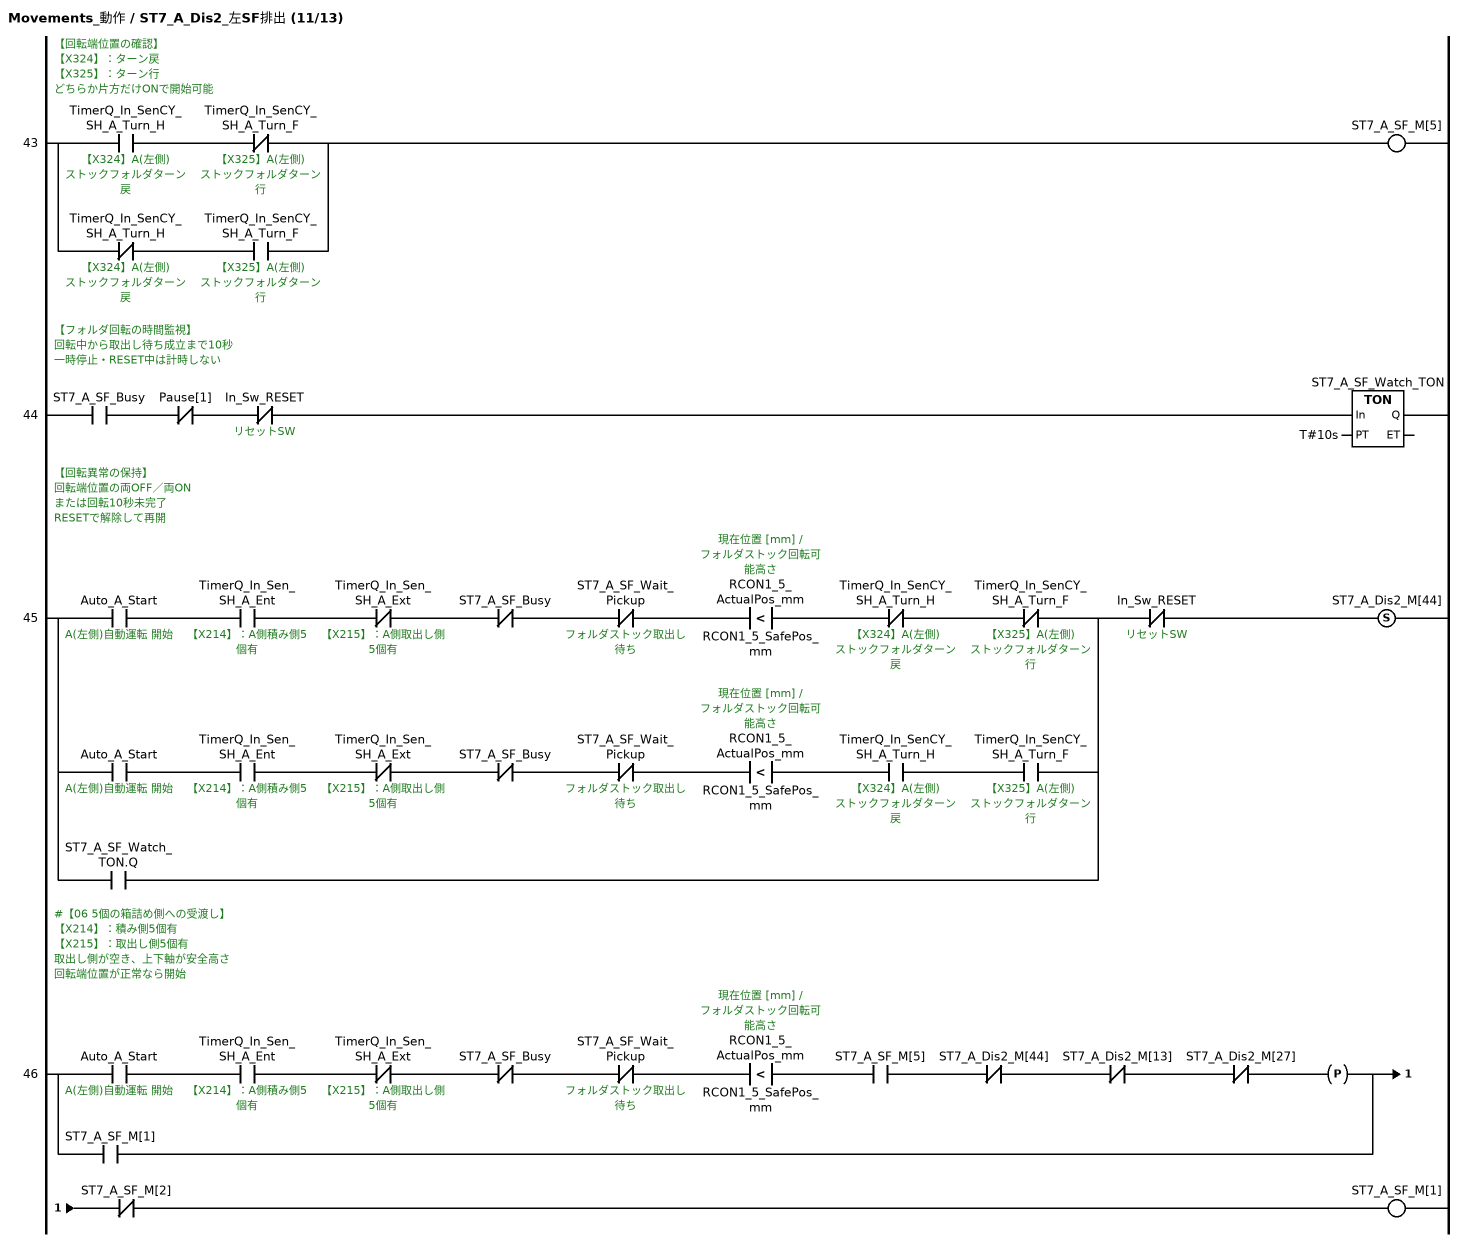
(* Rung 43: 【回転端位置の確認】 / 【X324】：ターン戻 / 【X325】：ターン行 / どちらか片方だけONで開始可能 *)
ST7_A_SF_M[5] := (TimerQ_In_SenCY_SH_A_Turn_H AND NOT TimerQ_In_SenCY_SH_A_Turn_F) OR (NOT TimerQ_In_SenCY_SH_A_Turn_H AND TimerQ_In_SenCY_SH_A_Turn_F);
(* Rung 44: 【フォルダ回転の時間監視】 / 回転中から取出し待ち成立まで10秒 / 一時停止・RESET中は計時しない *)
ST7_A_SF_Watch_TON(In := ST7_A_SF_Busy AND NOT Pause[1] AND NOT In_Sw_RESET, PT := T#10s);
(* Rung 45: 【回転異常の保持】 / 回転端位置の両OFF／両ON / または回転10秒未完了 / RESETで解除して再開 *)
IF ((Auto_A_Start AND TimerQ_In_Sen_SH_A_Ent AND NOT TimerQ_In_Sen_SH_A_Ext AND NOT ST7_A_SF_Busy AND NOT ST7_A_SF_Wait_Pickup AND (RCON1_5_ActualPos_mm < RCON1_5_SafePos_mm) AND NOT TimerQ_In_SenCY_SH_A_Turn_H AND NOT TimerQ_In_SenCY_SH_A_Turn_F) OR (Auto_A_Start AND TimerQ_In_Sen_SH_A_Ent AND NOT TimerQ_In_Sen_SH_A_Ext AND NOT ST7_A_SF_Busy AND NOT ST7_A_SF_Wait_Pickup AND (RCON1_5_ActualPos_mm < RCON1_5_SafePos_mm) AND TimerQ_In_SenCY_SH_A_Turn_H AND TimerQ_In_SenCY_SH_A_Turn_F) OR ST7_A_SF_Watch_TON.Q) AND NOT In_Sw_RESET THEN
    ST7_A_Dis2_M[44] := TRUE;
END_IF;
(* Rung 46: #【06 5個の箱詰め側への受渡し】 / 【X214】：積み側5個有 / 【X215】：取出し側5個有 / 取出し側が空き、上下軸が安全高さ / 回転端位置が正常なら開始 *)
_e112(CLK := Auto_A_Start AND TimerQ_In_Sen_SH_A_Ent AND NOT TimerQ_In_Sen_SH_A_Ext AND NOT ST7_A_SF_Busy AND NOT ST7_A_SF_Wait_Pickup AND (RCON1_5_ActualPos_mm < RCON1_5_SafePos_mm) AND ST7_A_SF_M[5] AND NOT ST7_A_Dis2_M[44] AND NOT ST7_A_Dis2_M[13] AND NOT ST7_A_Dis2_M[27]);
ST7_A_SF_M[1] := (_e112.Q OR ST7_A_SF_M[1]) AND NOT ST7_A_SF_M[2];

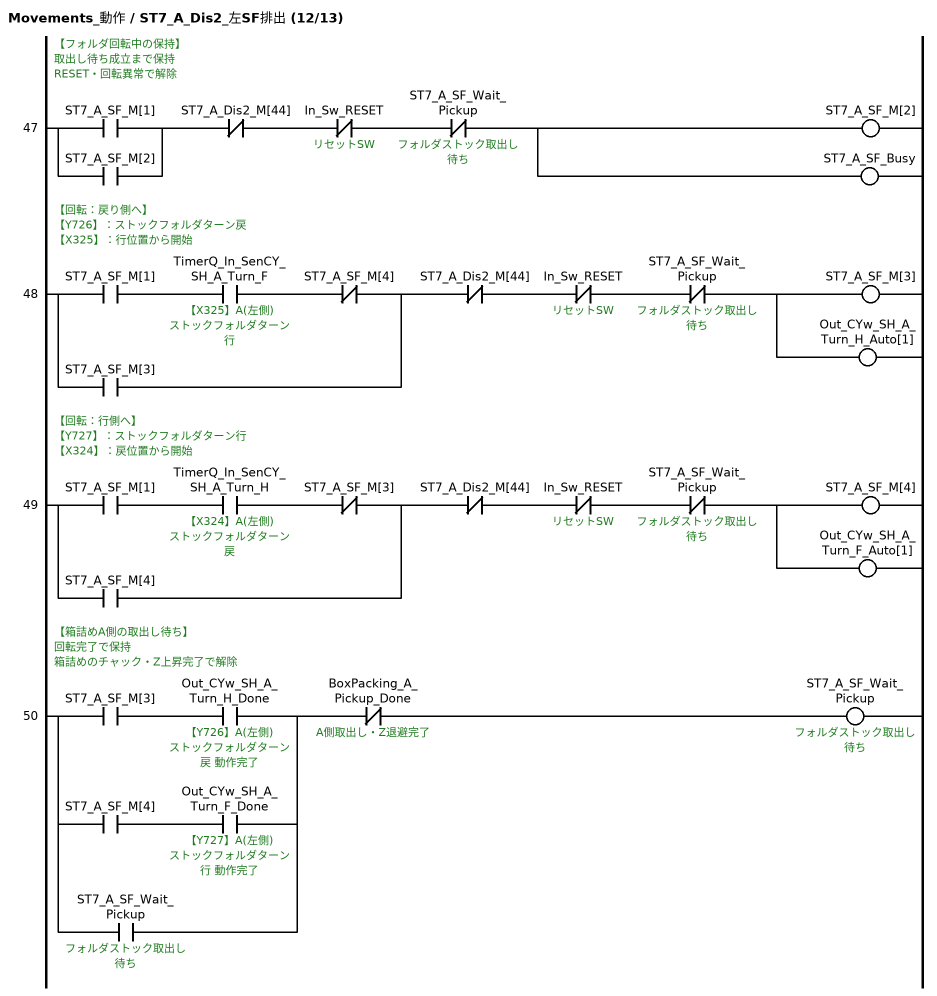
(* Rung 47: 【フォルダ回転中の保持】 / 取出し待ち成立まで保持 / RESET・回転異常で解除 *)
_p113 := (ST7_A_SF_M[1] OR ST7_A_SF_M[2]) AND NOT ST7_A_Dis2_M[44] AND NOT In_Sw_RESET AND NOT ST7_A_SF_Wait_Pickup;
ST7_A_SF_M[2] := _p113;
ST7_A_SF_Busy := _p113;
(* Rung 48: 【回転：戻り側へ】 / 【Y726】：ストックフォルダターン戻 / 【X325】：行位置から開始 *)
_p114 := ((ST7_A_SF_M[1] AND TimerQ_In_SenCY_SH_A_Turn_F AND NOT ST7_A_SF_M[4]) OR ST7_A_SF_M[3]) AND NOT ST7_A_Dis2_M[44] AND NOT In_Sw_RESET AND NOT ST7_A_SF_Wait_Pickup;
ST7_A_SF_M[3] := _p114;
Out_CYw_SH_A_Turn_H_Auto[1] := _p114;
(* Rung 49: 【回転：行側へ】 / 【Y727】：ストックフォルダターン行 / 【X324】：戻位置から開始 *)
_p115 := ((ST7_A_SF_M[1] AND TimerQ_In_SenCY_SH_A_Turn_H AND NOT ST7_A_SF_M[3]) OR ST7_A_SF_M[4]) AND NOT ST7_A_Dis2_M[44] AND NOT In_Sw_RESET AND NOT ST7_A_SF_Wait_Pickup;
ST7_A_SF_M[4] := _p115;
Out_CYw_SH_A_Turn_F_Auto[1] := _p115;
(* Rung 50: 【箱詰めA側の取出し待ち】 / 回転完了で保持 / 箱詰めのチャック・Z上昇完了で解除 *)
ST7_A_SF_Wait_Pickup := ((ST7_A_SF_M[3] AND Out_CYw_SH_A_Turn_H_Done) OR (ST7_A_SF_M[4] AND Out_CYw_SH_A_Turn_F_Done) OR ST7_A_SF_Wait_Pickup) AND NOT BoxPacking_A_Pickup_Done;

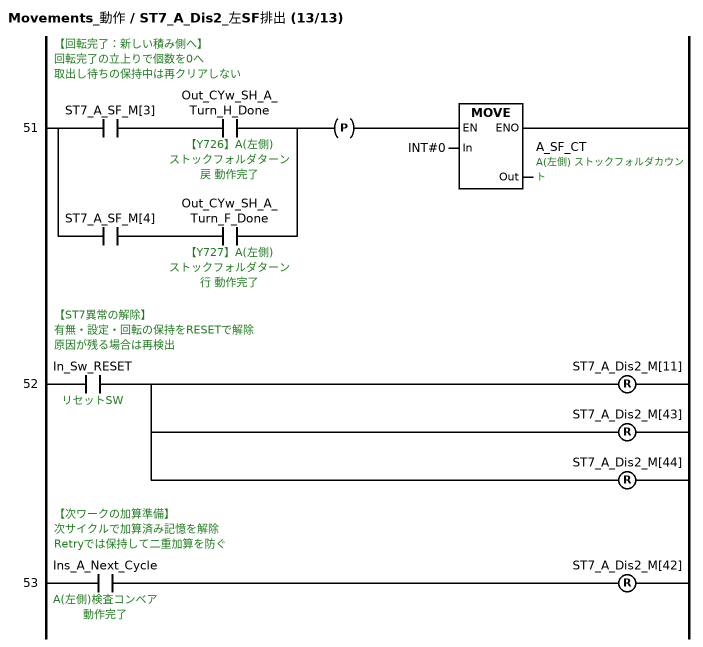
(* Rung 51: 【回転完了：新しい積み側へ】 / 回転完了の立上りで個数を0へ / 取出し待ちの保持中は再クリアしない *)
_e116(CLK := (ST7_A_SF_M[3] AND Out_CYw_SH_A_Turn_H_Done) OR (ST7_A_SF_M[4] AND Out_CYw_SH_A_Turn_F_Done));
IF _e116.Q THEN A_SF_CT := INT#0; END_IF;
(* Rung 52: 【ST7異常の解除】 / 有無・設定・回転の保持をRESETで解除 / 原因が残る場合は再検出 *)
IF In_Sw_RESET THEN
    ST7_A_Dis2_M[11] := FALSE;
    ST7_A_Dis2_M[43] := FALSE;
    ST7_A_Dis2_M[44] := FALSE;
END_IF;
(* Rung 53: 【次ワークの加算準備】 / 次サイクルで加算済み記憶を解除 / Retryでは保持して二重加算を防ぐ *)
IF Ins_A_Next_Cycle THEN ST7_A_Dis2_M[42] := FALSE; END_IF;

(* Section Destacker_段バラシ: ladder, written here as Structured Text *)

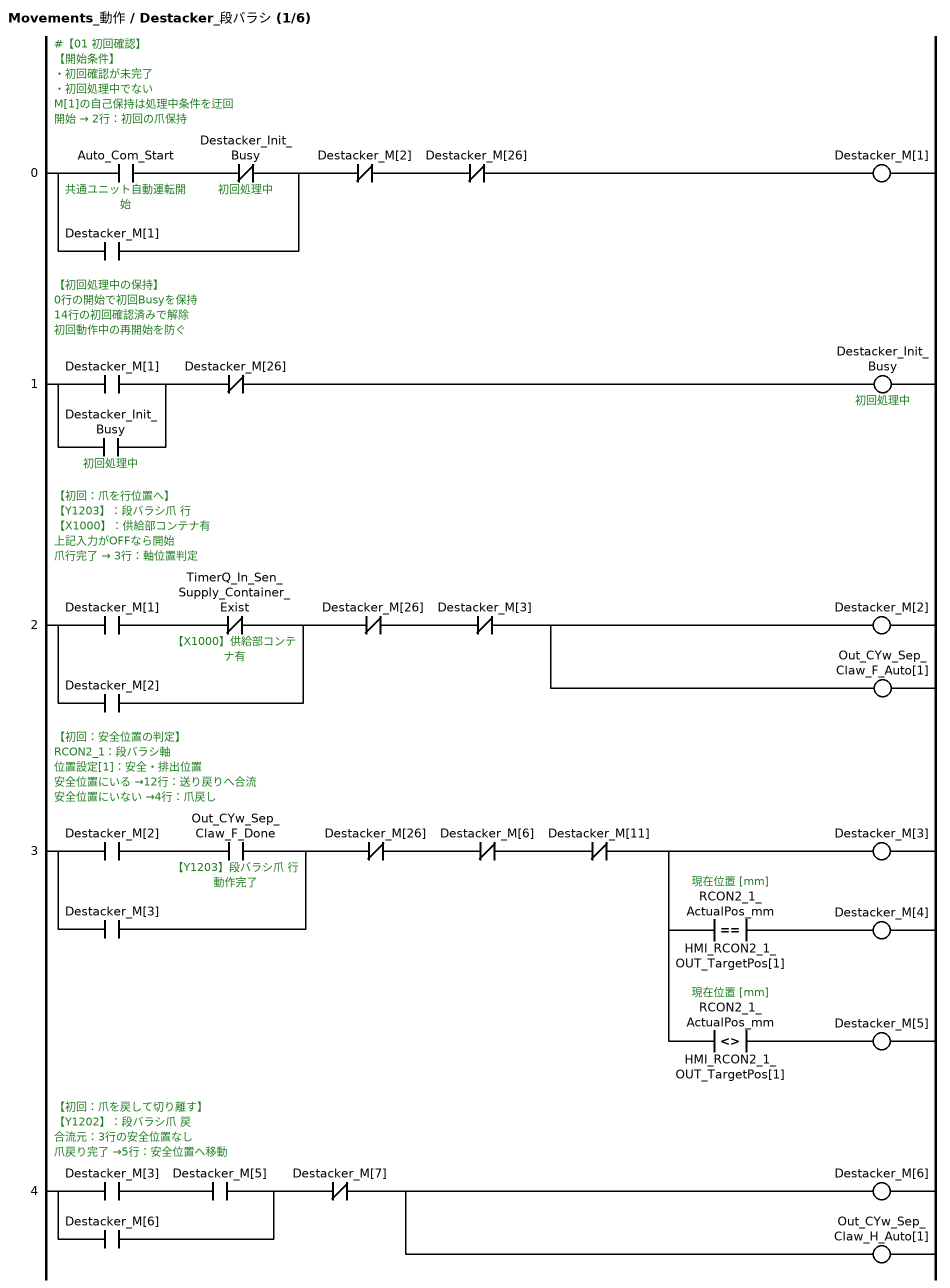
(* Rung 0: #【01 初回確認】 / 【開始条件】 / ・初回確認が未完了 / ・初回処理中でない / M[1]の自己保持は処理中条件を迂回 / 開始 → 2行：初回の爪保持 *)
Destacker_M[1] := ((Auto_Com_Start AND NOT Destacker_Init_Busy) OR Destacker_M[1]) AND NOT Destacker_M[2] AND NOT Destacker_M[26];
(* Rung 1: 【初回処理中の保持】 / 0行の開始で初回Busyを保持 / 14行の初回確認済みで解除 / 初回動作中の再開始を防ぐ *)
Destacker_Init_Busy := (Destacker_M[1] OR Destacker_Init_Busy) AND NOT Destacker_M[26];
(* Rung 2: 【初回：爪を行位置へ】 / 【Y1203】：段バラシ爪 行 / 【X1000】：供給部コンテナ有 / 上記入力がOFFなら開始 / 爪行完了 → 3行：軸位置判定 *)
_p117 := ((Destacker_M[1] AND NOT TimerQ_In_Sen_Supply_Container_Exist) OR Destacker_M[2]) AND NOT Destacker_M[26] AND NOT Destacker_M[3];
Destacker_M[2] := _p117;
Out_CYw_Sep_Claw_F_Auto[1] := _p117;
(* Rung 3: 【初回：安全位置の判定】 / RCON2_1：段バラシ軸 / 位置設定[1]：安全・排出位置 / 安全位置にいる →12行：送り戻りへ合流 / 安全位置にいない →4行：爪戻し *)
_p118 := ((Destacker_M[2] AND Out_CYw_Sep_Claw_F_Done) OR Destacker_M[3]) AND NOT Destacker_M[26] AND NOT Destacker_M[6] AND NOT Destacker_M[11];
Destacker_M[3] := _p118;
Destacker_M[4] := _p118 AND (RCON2_1_ActualPos_mm = HMI_RCON2_1_OUT_TargetPos[1]);
Destacker_M[5] := _p118 AND (RCON2_1_ActualPos_mm <> HMI_RCON2_1_OUT_TargetPos[1]);
(* Rung 4: 【初回：爪を戻して切り離す】 / 【Y1202】：段バラシ爪 戻 / 合流元：3行の安全位置なし / 爪戻り完了 →5行：安全位置へ移動 *)
_p119 := ((Destacker_M[3] AND Destacker_M[5]) OR Destacker_M[6]) AND NOT Destacker_M[7];
Destacker_M[6] := _p119;
Out_CYw_Sep_Claw_H_Auto[1] := _p119;

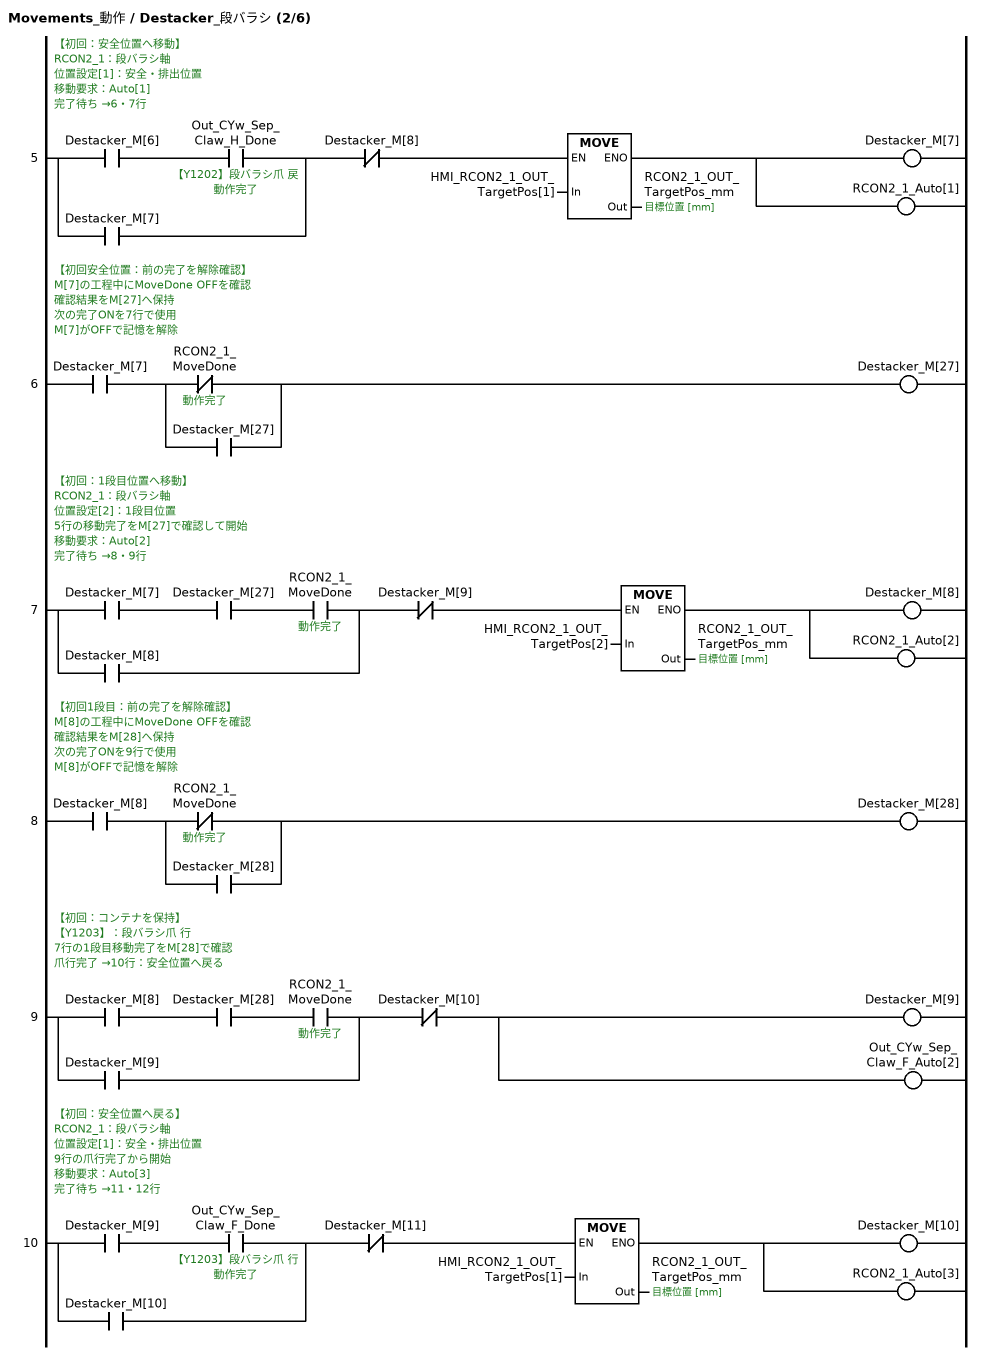
(* Rung 5: 【初回：安全位置へ移動】 / RCON2_1：段バラシ軸 / 位置設定[1]：安全・排出位置 / 移動要求：Auto[1] / 完了待ち →6・7行 *)
IF ((Destacker_M[6] AND Out_CYw_Sep_Claw_H_Done) OR Destacker_M[7]) AND NOT Destacker_M[8] THEN
    RCON2_1_OUT_TargetPos_mm := HMI_RCON2_1_OUT_TargetPos[1];
END_IF;
_p120 := ((Destacker_M[6] AND Out_CYw_Sep_Claw_H_Done) OR Destacker_M[7]) AND NOT Destacker_M[8];
Destacker_M[7] := _p120;
RCON2_1_Auto[1] := _p120;
(* Rung 6: 【初回安全位置：前の完了を解除確認】 / M[7]の工程中にMoveDone OFFを確認 / 確認結果をM[27]へ保持 / 次の完了ONを7行で使用 / M[7]がOFFで記憶を解除 *)
Destacker_M[27] := Destacker_M[7] AND (NOT RCON2_1_MoveDone OR Destacker_M[27]);
(* Rung 7: 【初回：1段目位置へ移動】 / RCON2_1：段バラシ軸 / 位置設定[2]：1段目位置 / 5行の移動完了をM[27]で確認して開始 / 移動要求：Auto[2] / 完了待ち →8・9行 *)
IF ((Destacker_M[7] AND Destacker_M[27] AND RCON2_1_MoveDone) OR Destacker_M[8]) AND NOT Destacker_M[9] THEN
    RCON2_1_OUT_TargetPos_mm := HMI_RCON2_1_OUT_TargetPos[2];
END_IF;
_p121 := ((Destacker_M[7] AND Destacker_M[27] AND RCON2_1_MoveDone) OR Destacker_M[8]) AND NOT Destacker_M[9];
Destacker_M[8] := _p121;
RCON2_1_Auto[2] := _p121;
(* Rung 8: 【初回1段目：前の完了を解除確認】 / M[8]の工程中にMoveDone OFFを確認 / 確認結果をM[28]へ保持 / 次の完了ONを9行で使用 / M[8]がOFFで記憶を解除 *)
Destacker_M[28] := Destacker_M[8] AND (NOT RCON2_1_MoveDone OR Destacker_M[28]);
(* Rung 9: 【初回：コンテナを保持】 / 【Y1203】：段バラシ爪 行 / 7行の1段目移動完了をM[28]で確認 / 爪行完了 →10行：安全位置へ戻る *)
_p122 := ((Destacker_M[8] AND Destacker_M[28] AND RCON2_1_MoveDone) OR Destacker_M[9]) AND NOT Destacker_M[10];
Destacker_M[9] := _p122;
Out_CYw_Sep_Claw_F_Auto[2] := _p122;
(* Rung 10: 【初回：安全位置へ戻る】 / RCON2_1：段バラシ軸 / 位置設定[1]：安全・排出位置 / 9行の爪行完了から開始 / 移動要求：Auto[3] / 完了待ち →11・12行 *)
IF ((Destacker_M[9] AND Out_CYw_Sep_Claw_F_Done) OR Destacker_M[10]) AND NOT Destacker_M[11] THEN
    RCON2_1_OUT_TargetPos_mm := HMI_RCON2_1_OUT_TargetPos[1];
END_IF;
_p123 := ((Destacker_M[9] AND Out_CYw_Sep_Claw_F_Done) OR Destacker_M[10]) AND NOT Destacker_M[11];
Destacker_M[10] := _p123;
RCON2_1_Auto[3] := _p123;

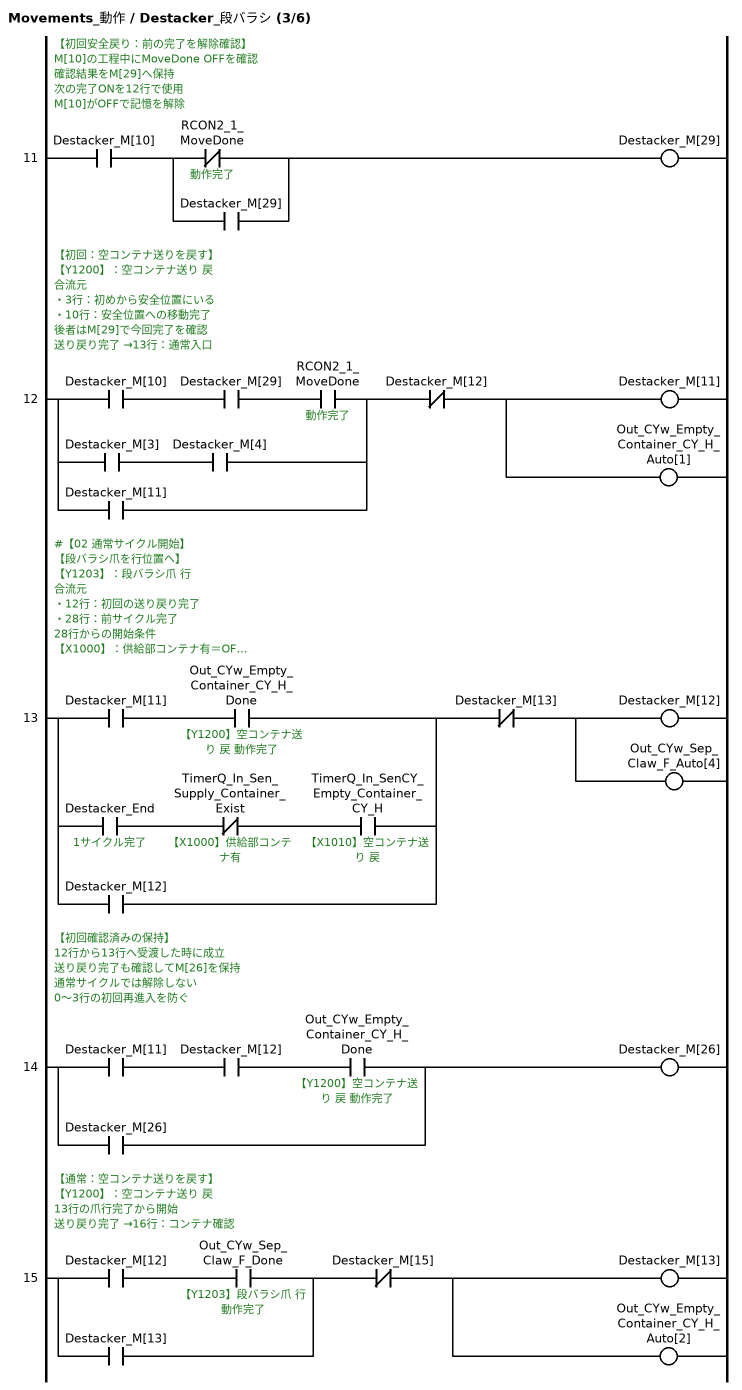
(* Rung 11: 【初回安全戻り：前の完了を解除確認】 / M[10]の工程中にMoveDone OFFを確認 / 確認結果をM[29]へ保持 / 次の完了ONを12行で使用 / M[10]がOFFで記憶を解除 *)
Destacker_M[29] := Destacker_M[10] AND (NOT RCON2_1_MoveDone OR Destacker_M[29]);
(* Rung 12: 【初回：空コンテナ送りを戻す】 / 【Y1200】：空コンテナ送り 戻 / 合流元 / ・3行：初めから安全位置にいる / ・10行：安全位置への移動完了 / 後者はM[29]で今回完了を確認 / 送り戻り完了 →13行：通常入口 *)
_p124 := ((Destacker_M[10] AND Destacker_M[29] AND RCON2_1_MoveDone) OR (Destacker_M[3] AND Destacker_M[4]) OR Destacker_M[11]) AND NOT Destacker_M[12];
Destacker_M[11] := _p124;
Out_CYw_Empty_Container_CY_H_Auto[1] := _p124;
(* Rung 13: #【02 通常サイクル開始】 / 【段バラシ爪を行位置へ】 / 【Y1203】：段バラシ爪 行 / 合流元 / ・12行：初回の送り戻り完了 / ・28行：前サイクル完了 / 28行からの開始条件 / 【X1000】：供給部コンテナ有＝OFF / 【X1010】：空コンテナ送り戻＝ON / 爪行完了 →15行：送り戻り確認 *)
_p125 := ((Destacker_M[11] AND Out_CYw_Empty_Container_CY_H_Done) OR (Destacker_End AND NOT TimerQ_In_Sen_Supply_Container_Exist AND TimerQ_In_SenCY_Empty_Container_CY_H) OR Destacker_M[12]) AND NOT Destacker_M[13];
Destacker_M[12] := _p125;
Out_CYw_Sep_Claw_F_Auto[4] := _p125;
(* Rung 14: 【初回確認済みの保持】 / 12行から13行へ受渡した時に成立 / 送り戻り完了も確認してM[26]を保持 / 通常サイクルでは解除しない / 0～3行の初回再進入を防ぐ *)
Destacker_M[26] := (Destacker_M[11] AND Destacker_M[12] AND Out_CYw_Empty_Container_CY_H_Done) OR Destacker_M[26];
(* Rung 15: 【通常：空コンテナ送りを戻す】 / 【Y1200】：空コンテナ送り 戻 / 13行の爪行完了から開始 / 送り戻り完了 →16行：コンテナ確認 *)
_p126 := ((Destacker_M[12] AND Out_CYw_Sep_Claw_F_Done) OR Destacker_M[13]) AND NOT Destacker_M[15];
Destacker_M[13] := _p126;
Out_CYw_Empty_Container_CY_H_Auto[2] := _p126;

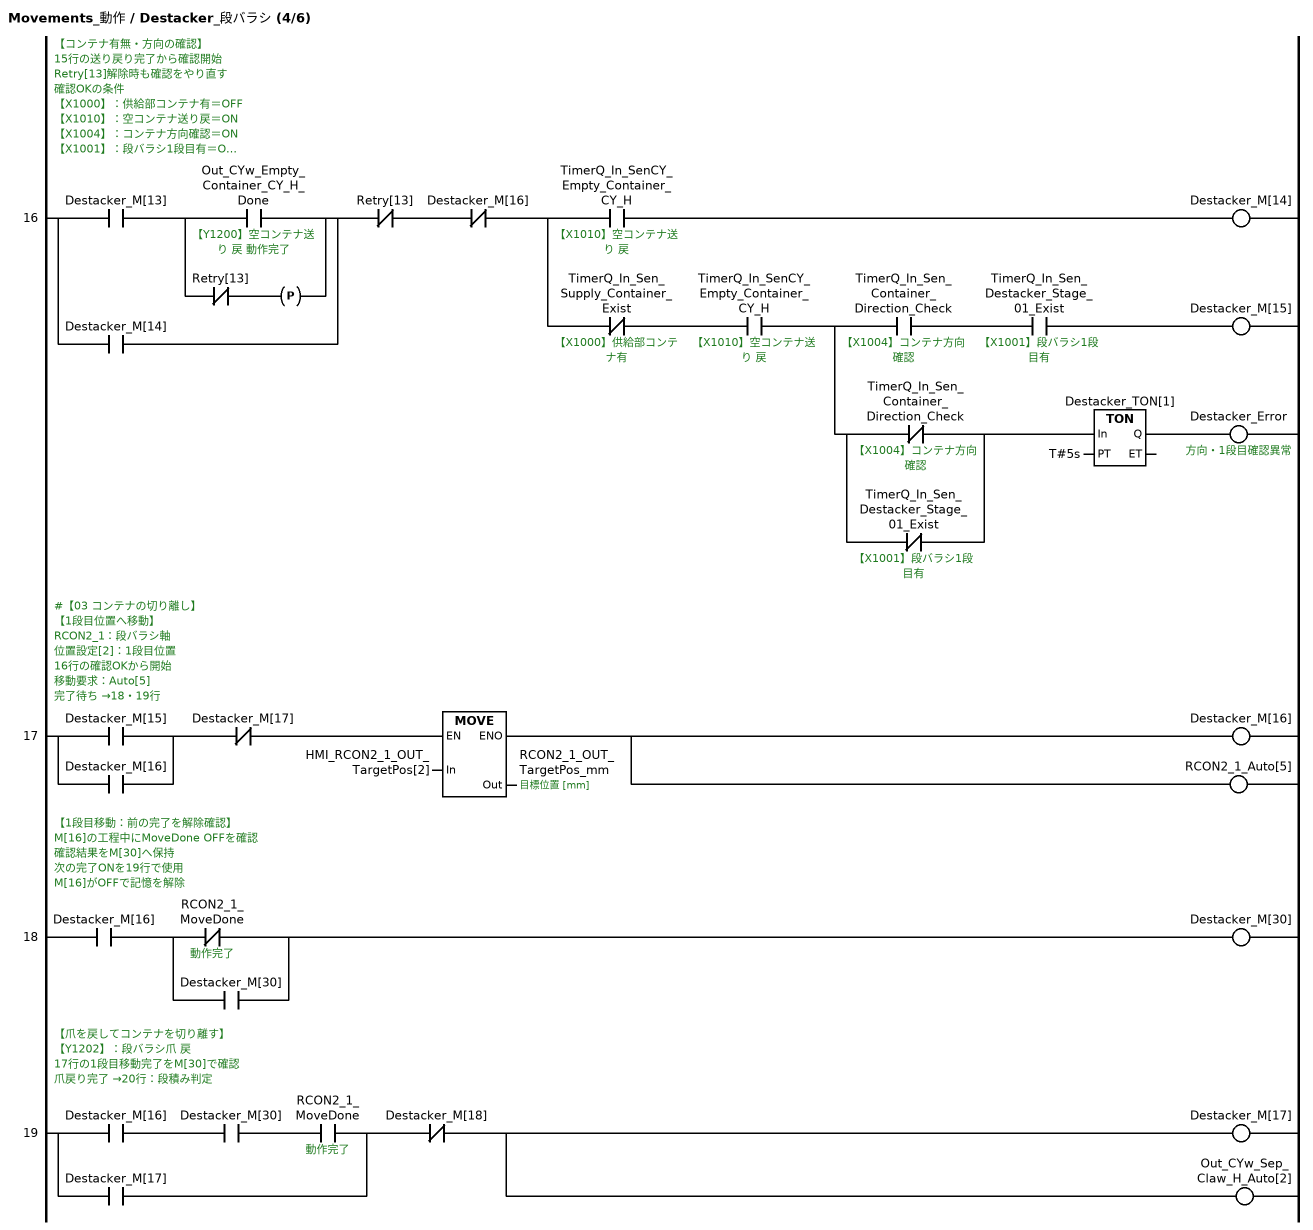
(* Rung 16: 【コンテナ有無・方向の確認】 / 15行の送り戻り完了から確認開始 / Retry[13]解除時も確認をやり直す / 確認OKの条件 / 【X1000】：供給部コンテナ有＝OFF / 【X1010】：空コンテナ送り戻＝ON / 【X1004】：コンテナ方向確認＝ON / 【X1001】：段バラシ1段目有＝ON / 確認OK →17行：1段目移動 / 方向NG／1段目なしが5秒 →確認異常 *)
_e127(CLK := Destacker_M[13] AND NOT Retry[13]);
_p128 := ((Destacker_M[13] AND Out_CYw_Empty_Container_CY_H_Done) OR _e127.Q OR Destacker_M[14]) AND NOT Retry[13] AND NOT Destacker_M[16];
Destacker_M[14] := _p128 AND TimerQ_In_SenCY_Empty_Container_CY_H;
_p129 := _p128 AND NOT TimerQ_In_Sen_Supply_Container_Exist AND TimerQ_In_SenCY_Empty_Container_CY_H;
Destacker_M[15] := _p129 AND TimerQ_In_Sen_Container_Direction_Check AND TimerQ_In_Sen_Destacker_Stage_01_Exist;
Destacker_TON[1](In := _p129 AND (NOT TimerQ_In_Sen_Container_Direction_Check OR NOT TimerQ_In_Sen_Destacker_Stage_01_Exist), PT := T#5s);
Destacker_Error := Destacker_TON[1].Q;
(* Rung 17: #【03 コンテナの切り離し】 / 【1段目位置へ移動】 / RCON2_1：段バラシ軸 / 位置設定[2]：1段目位置 / 16行の確認OKから開始 / 移動要求：Auto[5] / 完了待ち →18・19行 *)
IF (Destacker_M[15] OR Destacker_M[16]) AND NOT Destacker_M[17] THEN
    RCON2_1_OUT_TargetPos_mm := HMI_RCON2_1_OUT_TargetPos[2];
END_IF;
_p130 := (Destacker_M[15] OR Destacker_M[16]) AND NOT Destacker_M[17];
Destacker_M[16] := _p130;
RCON2_1_Auto[5] := _p130;
(* Rung 18: 【1段目移動：前の完了を解除確認】 / M[16]の工程中にMoveDone OFFを確認 / 確認結果をM[30]へ保持 / 次の完了ONを19行で使用 / M[16]がOFFで記憶を解除 *)
Destacker_M[30] := Destacker_M[16] AND (NOT RCON2_1_MoveDone OR Destacker_M[30]);
(* Rung 19: 【爪を戻してコンテナを切り離す】 / 【Y1202】：段バラシ爪 戻 / 17行の1段目移動完了をM[30]で確認 / 爪戻り完了 →20行：段積み判定 *)
_p131 := ((Destacker_M[16] AND Destacker_M[30] AND RCON2_1_MoveDone) OR Destacker_M[17]) AND NOT Destacker_M[18];
Destacker_M[17] := _p131;
Out_CYw_Sep_Claw_H_Auto[2] := _p131;

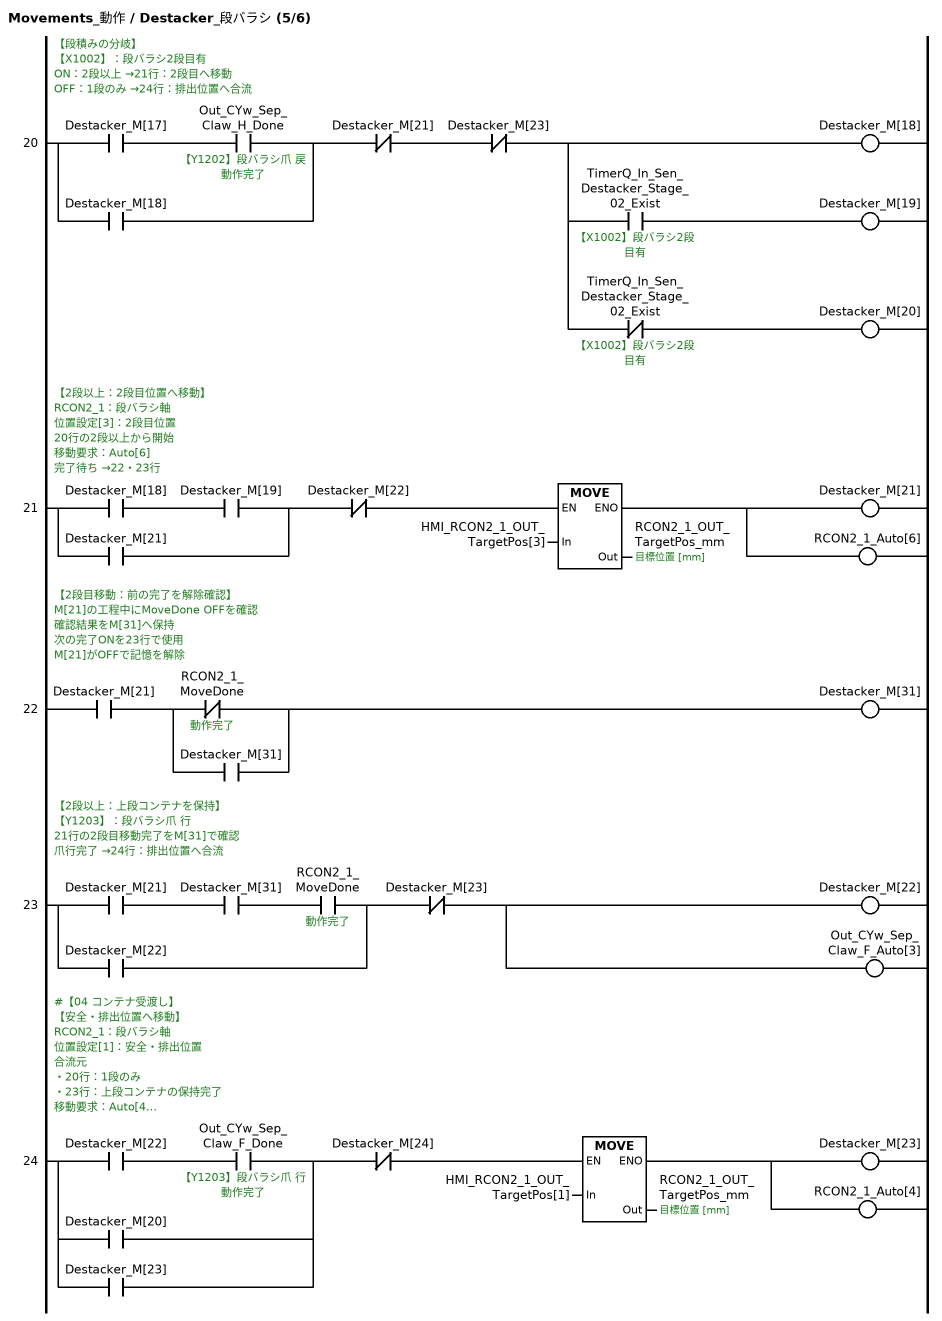
(* Rung 20: 【段積みの分岐】 / 【X1002】：段バラシ2段目有 / ON：2段以上 →21行：2段目へ移動 / OFF：1段のみ →24行：排出位置へ合流 *)
_p132 := ((Destacker_M[17] AND Out_CYw_Sep_Claw_H_Done) OR Destacker_M[18]) AND NOT Destacker_M[21] AND NOT Destacker_M[23];
Destacker_M[18] := _p132;
Destacker_M[19] := _p132 AND TimerQ_In_Sen_Destacker_Stage_02_Exist;
Destacker_M[20] := _p132 AND NOT TimerQ_In_Sen_Destacker_Stage_02_Exist;
(* Rung 21: 【2段以上：2段目位置へ移動】 / RCON2_1：段バラシ軸 / 位置設定[3]：2段目位置 / 20行の2段以上から開始 / 移動要求：Auto[6] / 完了待ち →22・23行 *)
IF ((Destacker_M[18] AND Destacker_M[19]) OR Destacker_M[21]) AND NOT Destacker_M[22] THEN
    RCON2_1_OUT_TargetPos_mm := HMI_RCON2_1_OUT_TargetPos[3];
END_IF;
_p133 := ((Destacker_M[18] AND Destacker_M[19]) OR Destacker_M[21]) AND NOT Destacker_M[22];
Destacker_M[21] := _p133;
RCON2_1_Auto[6] := _p133;
(* Rung 22: 【2段目移動：前の完了を解除確認】 / M[21]の工程中にMoveDone OFFを確認 / 確認結果をM[31]へ保持 / 次の完了ONを23行で使用 / M[21]がOFFで記憶を解除 *)
Destacker_M[31] := Destacker_M[21] AND (NOT RCON2_1_MoveDone OR Destacker_M[31]);
(* Rung 23: 【2段以上：上段コンテナを保持】 / 【Y1203】：段バラシ爪 行 / 21行の2段目移動完了をM[31]で確認 / 爪行完了 →24行：排出位置へ合流 *)
_p134 := ((Destacker_M[21] AND Destacker_M[31] AND RCON2_1_MoveDone) OR Destacker_M[22]) AND NOT Destacker_M[23];
Destacker_M[22] := _p134;
Out_CYw_Sep_Claw_F_Auto[3] := _p134;
(* Rung 24: #【04 コンテナ受渡し】 / 【安全・排出位置へ移動】 / RCON2_1：段バラシ軸 / 位置設定[1]：安全・排出位置 / 合流元 / ・20行：1段のみ / ・23行：上段コンテナの保持完了 / 移動要求：Auto[4] / 完了待ち →25・26行 *)
IF ((Destacker_M[22] AND Out_CYw_Sep_Claw_F_Done) OR Destacker_M[20] OR Destacker_M[23]) AND NOT Destacker_M[24] THEN
    RCON2_1_OUT_TargetPos_mm := HMI_RCON2_1_OUT_TargetPos[1];
END_IF;
_p135 := ((Destacker_M[22] AND Out_CYw_Sep_Claw_F_Done) OR Destacker_M[20] OR Destacker_M[23]) AND NOT Destacker_M[24];
Destacker_M[23] := _p135;
RCON2_1_Auto[4] := _p135;

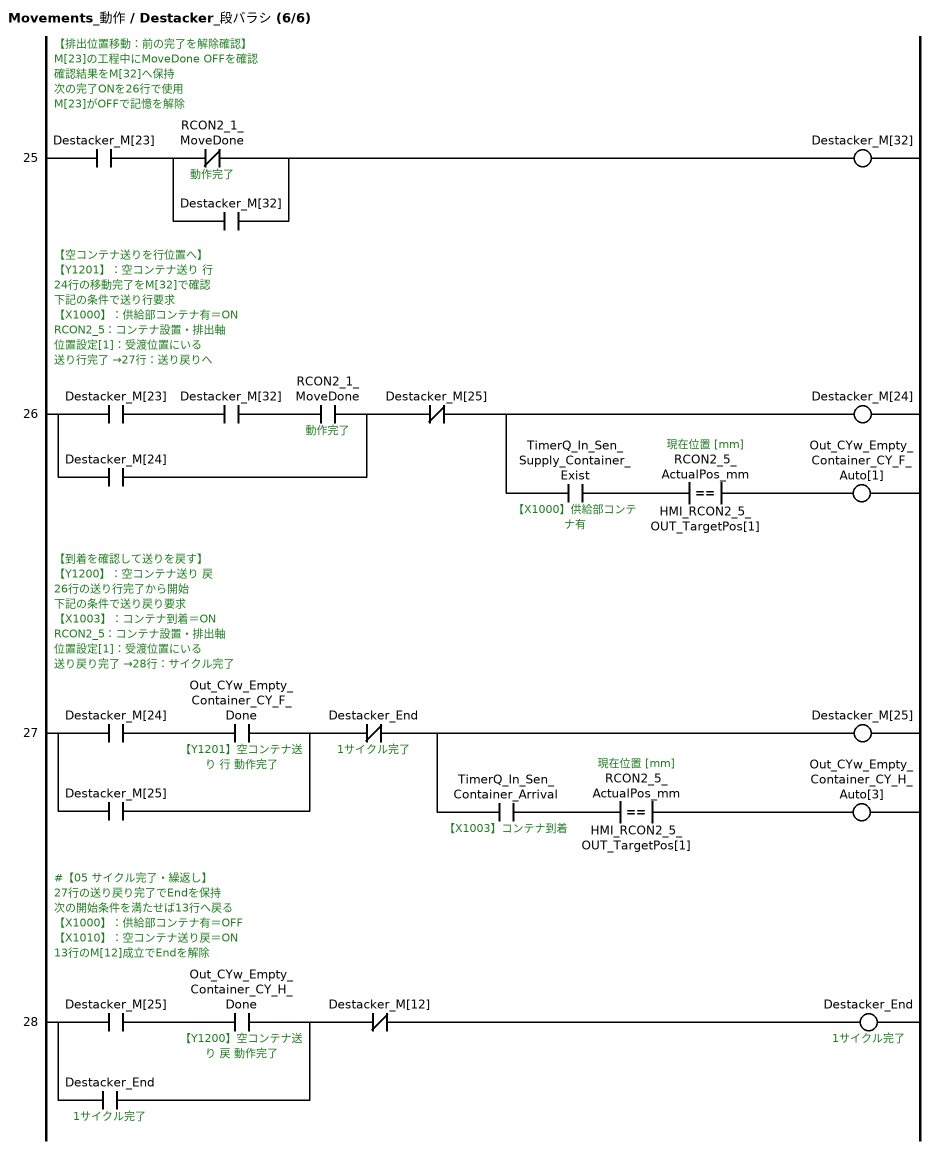
(* Rung 25: 【排出位置移動：前の完了を解除確認】 / M[23]の工程中にMoveDone OFFを確認 / 確認結果をM[32]へ保持 / 次の完了ONを26行で使用 / M[23]がOFFで記憶を解除 *)
Destacker_M[32] := Destacker_M[23] AND (NOT RCON2_1_MoveDone OR Destacker_M[32]);
(* Rung 26: 【空コンテナ送りを行位置へ】 / 【Y1201】：空コンテナ送り 行 / 24行の移動完了をM[32]で確認 / 下記の条件で送り行要求 / 【X1000】：供給部コンテナ有＝ON / RCON2_5：コンテナ設置・排出軸 / 位置設定[1]：受渡位置にいる / 送り行完了 →27行：送り戻りへ *)
_p136 := ((Destacker_M[23] AND Destacker_M[32] AND RCON2_1_MoveDone) OR Destacker_M[24]) AND NOT Destacker_M[25];
Destacker_M[24] := _p136;
Out_CYw_Empty_Container_CY_F_Auto[1] := _p136 AND TimerQ_In_Sen_Supply_Container_Exist AND (RCON2_5_ActualPos_mm = HMI_RCON2_5_OUT_TargetPos[1]);
(* Rung 27: 【到着を確認して送りを戻す】 / 【Y1200】：空コンテナ送り 戻 / 26行の送り行完了から開始 / 下記の条件で送り戻り要求 / 【X1003】：コンテナ到着＝ON / RCON2_5：コンテナ設置・排出軸 / 位置設定[1]：受渡位置にいる / 送り戻り完了 →28行：サイクル完了 *)
_p137 := ((Destacker_M[24] AND Out_CYw_Empty_Container_CY_F_Done) OR Destacker_M[25]) AND NOT Destacker_End;
Destacker_M[25] := _p137;
Out_CYw_Empty_Container_CY_H_Auto[3] := _p137 AND TimerQ_In_Sen_Container_Arrival AND (RCON2_5_ActualPos_mm = HMI_RCON2_5_OUT_TargetPos[1]);
(* Rung 28: #【05 サイクル完了・繰返し】 / 27行の送り戻り完了でEndを保持 / 次の開始条件を満たせば13行へ戻る / 【X1000】：供給部コンテナ有＝OFF / 【X1010】：空コンテナ送り戻＝ON / 13行のM[12]成立でEndを解除 *)
Destacker_End := ((Destacker_M[25] AND Out_CYw_Empty_Container_CY_H_Done) OR Destacker_End) AND NOT Destacker_M[12];

(* Section BoxPacking_箱詰め: ladder, written here as Structured Text *)

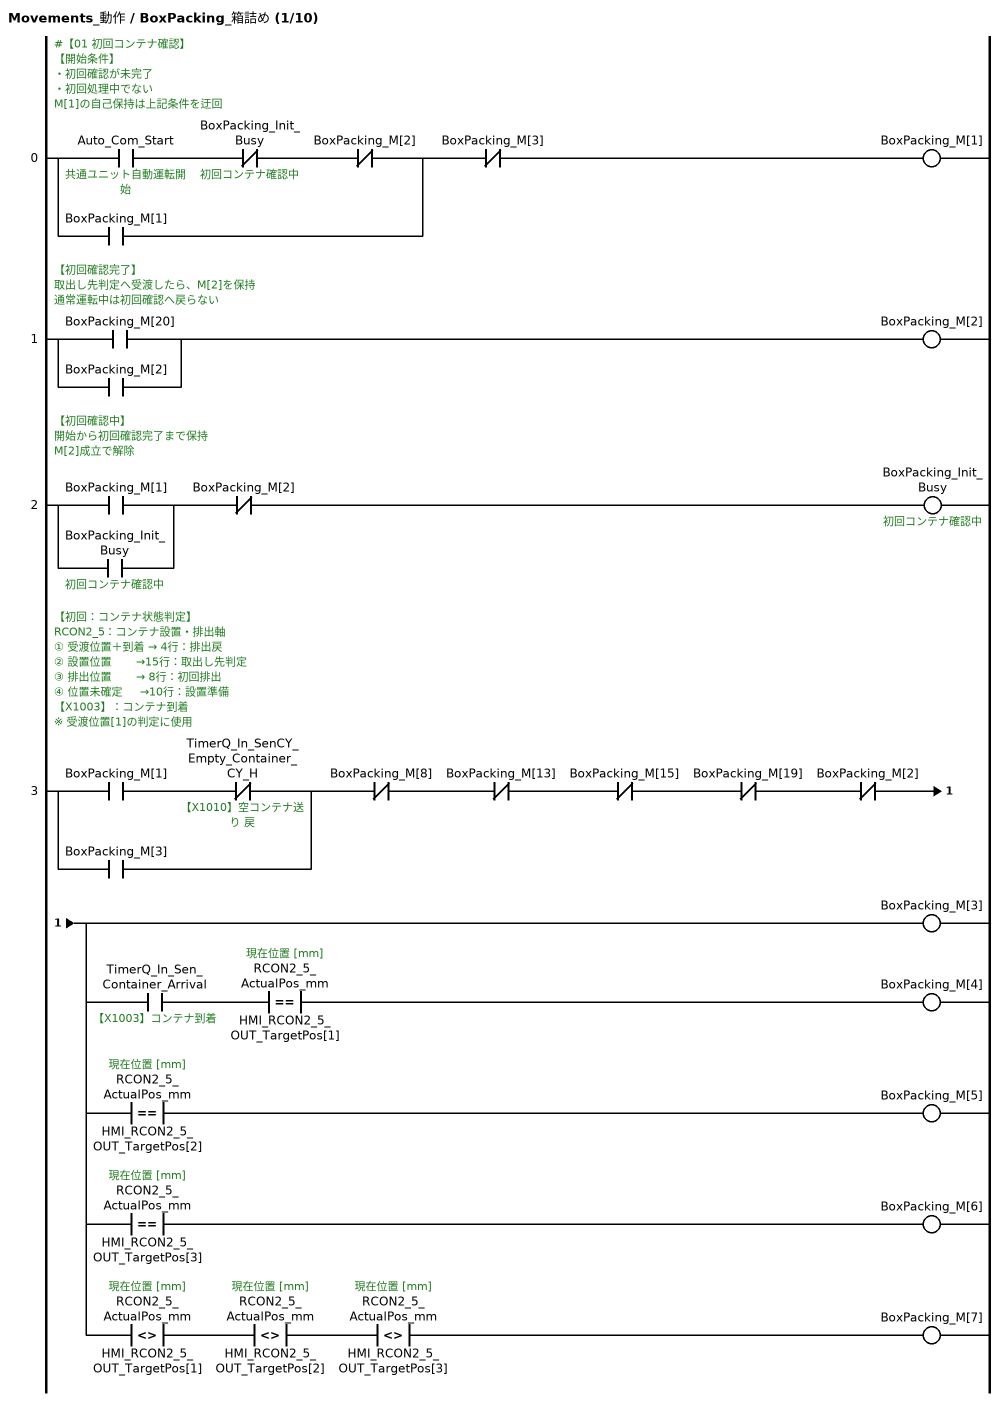
(* Rung 0: #【01 初回コンテナ確認】 / 【開始条件】 / ・初回確認が未完了 / ・初回処理中でない / M[1]の自己保持は上記条件を迂回 *)
BoxPacking_M[1] := ((Auto_Com_Start AND NOT BoxPacking_Init_Busy AND NOT BoxPacking_M[2]) OR BoxPacking_M[1]) AND NOT BoxPacking_M[3];
(* Rung 1: 【初回確認完了】 / 取出し先判定へ受渡したら、M[2]を保持 / 通常運転中は初回確認へ戻らない *)
BoxPacking_M[2] := BoxPacking_M[20] OR BoxPacking_M[2];
(* Rung 2: 【初回確認中】 / 開始から初回確認完了まで保持 / M[2]成立で解除 *)
BoxPacking_Init_Busy := (BoxPacking_M[1] OR BoxPacking_Init_Busy) AND NOT BoxPacking_M[2];
(* Rung 3: 【初回：コンテナ状態判定】 / RCON2_5：コンテナ設置・排出軸 / ① 受渡位置＋到着 → 4行：排出戻 / ② 設置位置       →15行：取出し先判定 / ③ 排出位置       → 8行：初回排出 / ④ 位置未確定     →10行：設置準備 / 【X1003】：コンテナ到着 / ※ 受渡位置[1]の判定に使用 *)
_p138 := ((BoxPacking_M[1] AND NOT TimerQ_In_SenCY_Empty_Container_CY_H) OR BoxPacking_M[3]) AND NOT BoxPacking_M[8] AND NOT BoxPacking_M[13] AND NOT BoxPacking_M[15] AND NOT BoxPacking_M[19] AND NOT BoxPacking_M[2];
BoxPacking_M[3] := _p138;
BoxPacking_M[4] := _p138 AND TimerQ_In_Sen_Container_Arrival AND (RCON2_5_ActualPos_mm = HMI_RCON2_5_OUT_TargetPos[1]);
BoxPacking_M[5] := _p138 AND (RCON2_5_ActualPos_mm = HMI_RCON2_5_OUT_TargetPos[2]);
BoxPacking_M[6] := _p138 AND (RCON2_5_ActualPos_mm = HMI_RCON2_5_OUT_TargetPos[3]);
BoxPacking_M[7] := _p138 AND (RCON2_5_ActualPos_mm <> HMI_RCON2_5_OUT_TargetPos[1]) AND (RCON2_5_ActualPos_mm <> HMI_RCON2_5_OUT_TargetPos[2]) AND (RCON2_5_ActualPos_mm <> HMI_RCON2_5_OUT_TargetPos[3]);

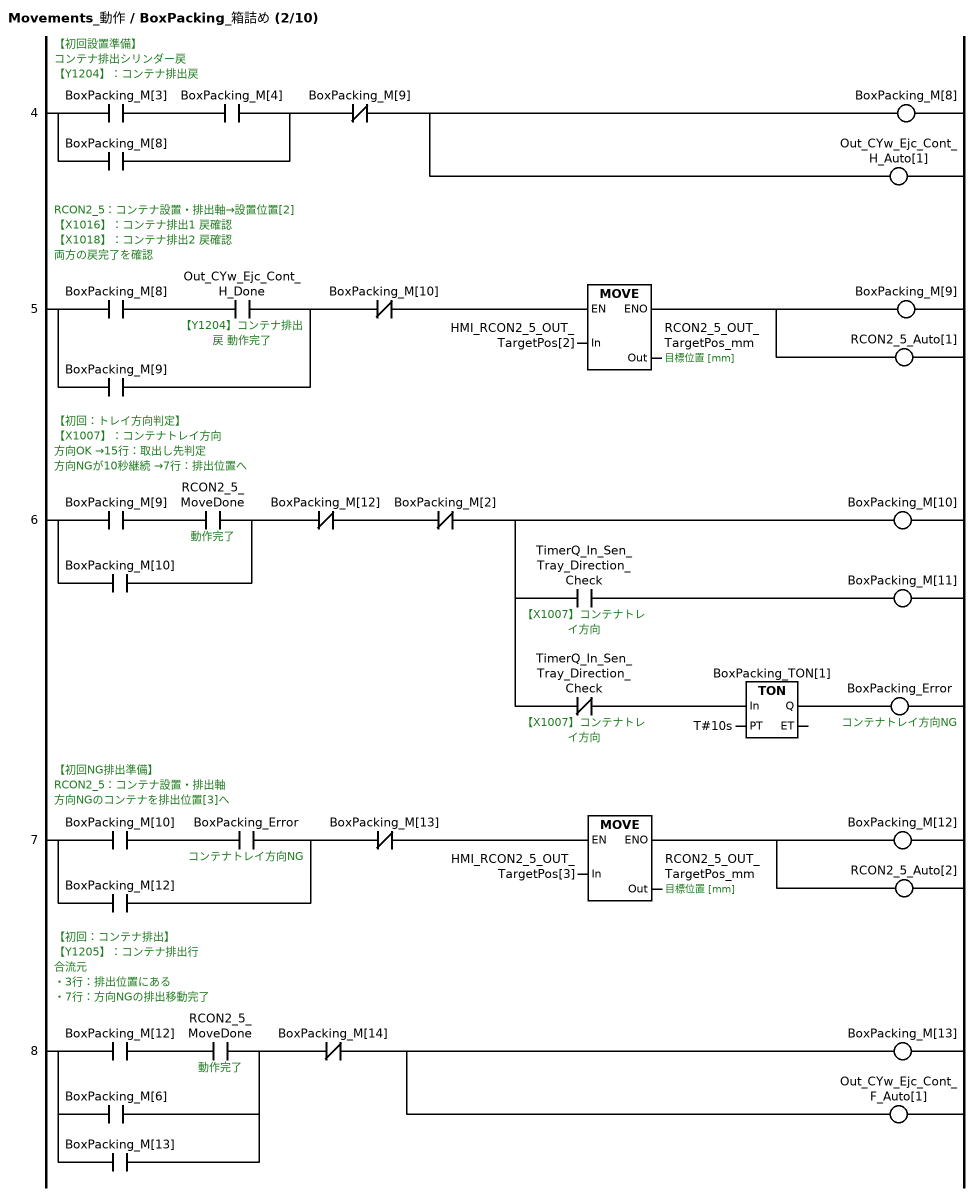
(* Rung 4: 【初回設置準備】 / コンテナ排出シリンダー戻 / 【Y1204】：コンテナ排出戻 *)
_p139 := ((BoxPacking_M[3] AND BoxPacking_M[4]) OR BoxPacking_M[8]) AND NOT BoxPacking_M[9];
BoxPacking_M[8] := _p139;
Out_CYw_Ejc_Cont_H_Auto[1] := _p139;
(* Rung 5: RCON2_5：コンテナ設置・排出軸→設置位置[2] / 【X1016】：コンテナ排出1 戻確認 / 【X1018】：コンテナ排出2 戻確認 / 両方の戻完了を確認 *)
IF ((BoxPacking_M[8] AND Out_CYw_Ejc_Cont_H_Done) OR BoxPacking_M[9]) AND NOT BoxPacking_M[10] THEN
    RCON2_5_OUT_TargetPos_mm := HMI_RCON2_5_OUT_TargetPos[2];
END_IF;
_p140 := ((BoxPacking_M[8] AND Out_CYw_Ejc_Cont_H_Done) OR BoxPacking_M[9]) AND NOT BoxPacking_M[10];
BoxPacking_M[9] := _p140;
RCON2_5_Auto[1] := _p140;
(* Rung 6: 【初回：トレイ方向判定】 / 【X1007】：コンテナトレイ方向 / 方向OK →15行：取出し先判定 / 方向NGが10秒継続 →7行：排出位置へ *)
_p141 := ((BoxPacking_M[9] AND RCON2_5_MoveDone) OR BoxPacking_M[10]) AND NOT BoxPacking_M[12] AND NOT BoxPacking_M[2];
BoxPacking_M[10] := _p141;
BoxPacking_M[11] := _p141 AND TimerQ_In_Sen_Tray_Direction_Check;
BoxPacking_TON[1](In := _p141 AND NOT TimerQ_In_Sen_Tray_Direction_Check, PT := T#10s);
BoxPacking_Error := BoxPacking_TON[1].Q;
(* Rung 7: 【初回NG排出準備】 / RCON2_5：コンテナ設置・排出軸 / 方向NGのコンテナを排出位置[3]へ *)
IF ((BoxPacking_M[10] AND BoxPacking_Error) OR BoxPacking_M[12]) AND NOT BoxPacking_M[13] THEN
    RCON2_5_OUT_TargetPos_mm := HMI_RCON2_5_OUT_TargetPos[3];
END_IF;
_p142 := ((BoxPacking_M[10] AND BoxPacking_Error) OR BoxPacking_M[12]) AND NOT BoxPacking_M[13];
BoxPacking_M[12] := _p142;
RCON2_5_Auto[2] := _p142;
(* Rung 8: 【初回：コンテナ排出】 / 【Y1205】：コンテナ排出行 / 合流元 / ・3行：排出位置にある / ・7行：方向NGの排出移動完了 *)
_p143 := ((BoxPacking_M[12] AND RCON2_5_MoveDone) OR BoxPacking_M[6] OR BoxPacking_M[13]) AND NOT BoxPacking_M[14];
BoxPacking_M[13] := _p143;
Out_CYw_Ejc_Cont_F_Auto[1] := _p143;

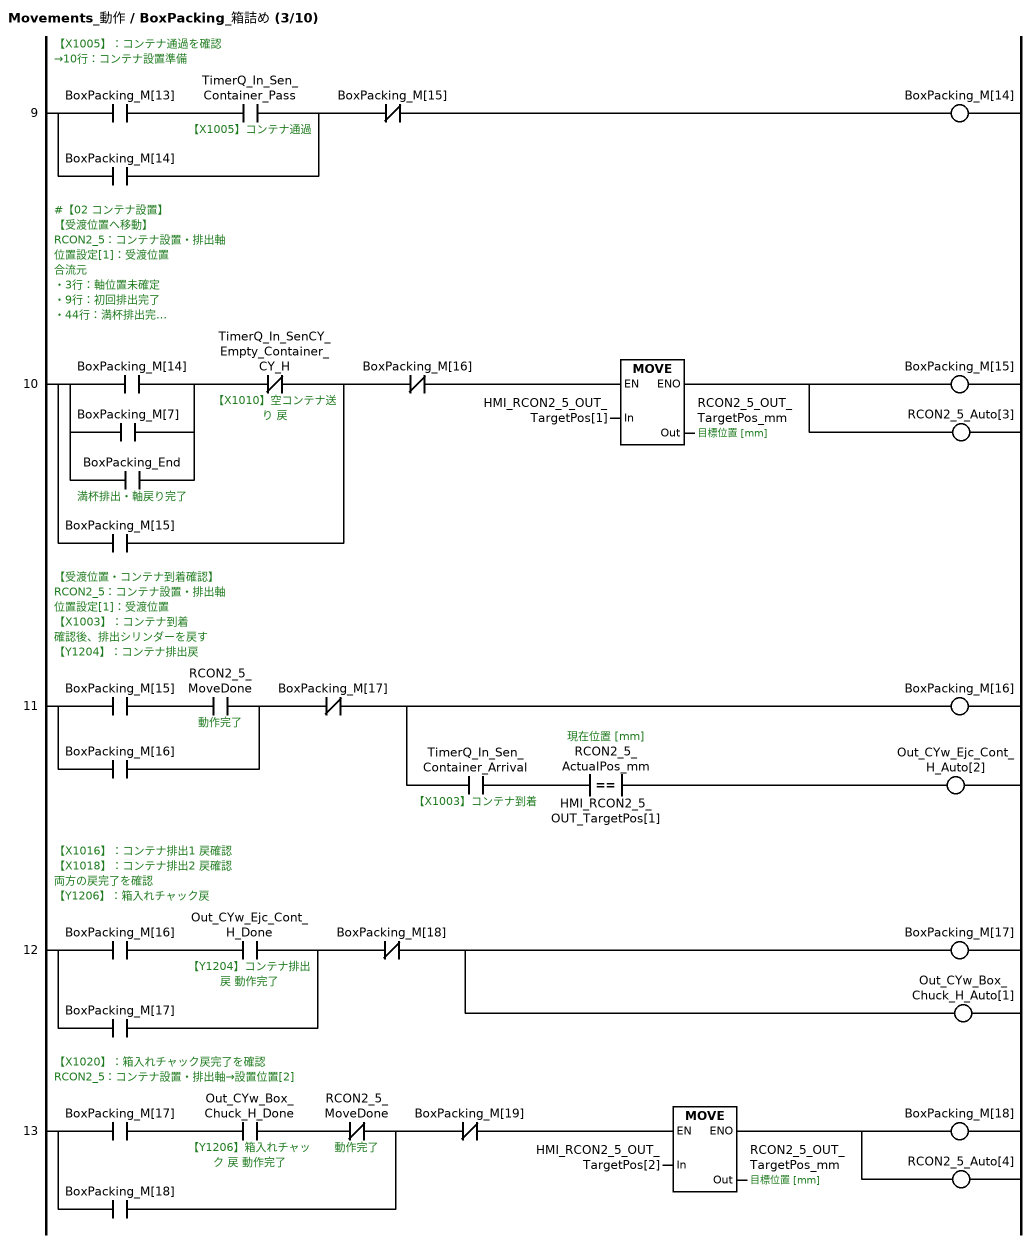
(* Rung 9: 【X1005】：コンテナ通過を確認 / →10行：コンテナ設置準備 *)
BoxPacking_M[14] := ((BoxPacking_M[13] AND TimerQ_In_Sen_Container_Pass) OR BoxPacking_M[14]) AND NOT BoxPacking_M[15];
(* Rung 10: #【02 コンテナ設置】 / 【受渡位置へ移動】 / RCON2_5：コンテナ設置・排出軸 / 位置設定[1]：受渡位置 / 合流元 / ・3行：軸位置未確定 / ・9行：初回排出完了 / ・44行：満杯排出完了 / 44行からは、下記入力のOFFで復帰 / 【X1010】：空コンテナ送り戻確認 *)
IF (((BoxPacking_M[14] OR BoxPacking_M[7] OR BoxPacking_End) AND NOT TimerQ_In_SenCY_Empty_Container_CY_H) OR BoxPacking_M[15]) AND NOT BoxPacking_M[16] THEN
    RCON2_5_OUT_TargetPos_mm := HMI_RCON2_5_OUT_TargetPos[1];
END_IF;
_p144 := (((BoxPacking_M[14] OR BoxPacking_M[7] OR BoxPacking_End) AND NOT TimerQ_In_SenCY_Empty_Container_CY_H) OR BoxPacking_M[15]) AND NOT BoxPacking_M[16];
BoxPacking_M[15] := _p144;
RCON2_5_Auto[3] := _p144;
(* Rung 11: 【受渡位置・コンテナ到着確認】 / RCON2_5：コンテナ設置・排出軸 / 位置設定[1]：受渡位置 / 【X1003】：コンテナ到着 / 確認後、排出シリンダーを戻す / 【Y1204】：コンテナ排出戻 *)
_p145 := ((BoxPacking_M[15] AND RCON2_5_MoveDone) OR BoxPacking_M[16]) AND NOT BoxPacking_M[17];
BoxPacking_M[16] := _p145;
Out_CYw_Ejc_Cont_H_Auto[2] := _p145 AND TimerQ_In_Sen_Container_Arrival AND (RCON2_5_ActualPos_mm = HMI_RCON2_5_OUT_TargetPos[1]);
(* Rung 12: 【X1016】：コンテナ排出1 戻確認 / 【X1018】：コンテナ排出2 戻確認 / 両方の戻完了を確認 / 【Y1206】：箱入れチャック戻 *)
_p146 := ((BoxPacking_M[16] AND Out_CYw_Ejc_Cont_H_Done) OR BoxPacking_M[17]) AND NOT BoxPacking_M[18];
BoxPacking_M[17] := _p146;
Out_CYw_Box_Chuck_H_Auto[1] := _p146;
(* Rung 13: 【X1020】：箱入れチャック戻完了を確認 / RCON2_5：コンテナ設置・排出軸→設置位置[2] *)
IF ((BoxPacking_M[17] AND Out_CYw_Box_Chuck_H_Done AND NOT RCON2_5_MoveDone) OR BoxPacking_M[18]) AND NOT BoxPacking_M[19] THEN
    RCON2_5_OUT_TargetPos_mm := HMI_RCON2_5_OUT_TargetPos[2];
END_IF;
_p147 := ((BoxPacking_M[17] AND Out_CYw_Box_Chuck_H_Done AND NOT RCON2_5_MoveDone) OR BoxPacking_M[18]) AND NOT BoxPacking_M[19];
BoxPacking_M[18] := _p147;
RCON2_5_Auto[4] := _p147;

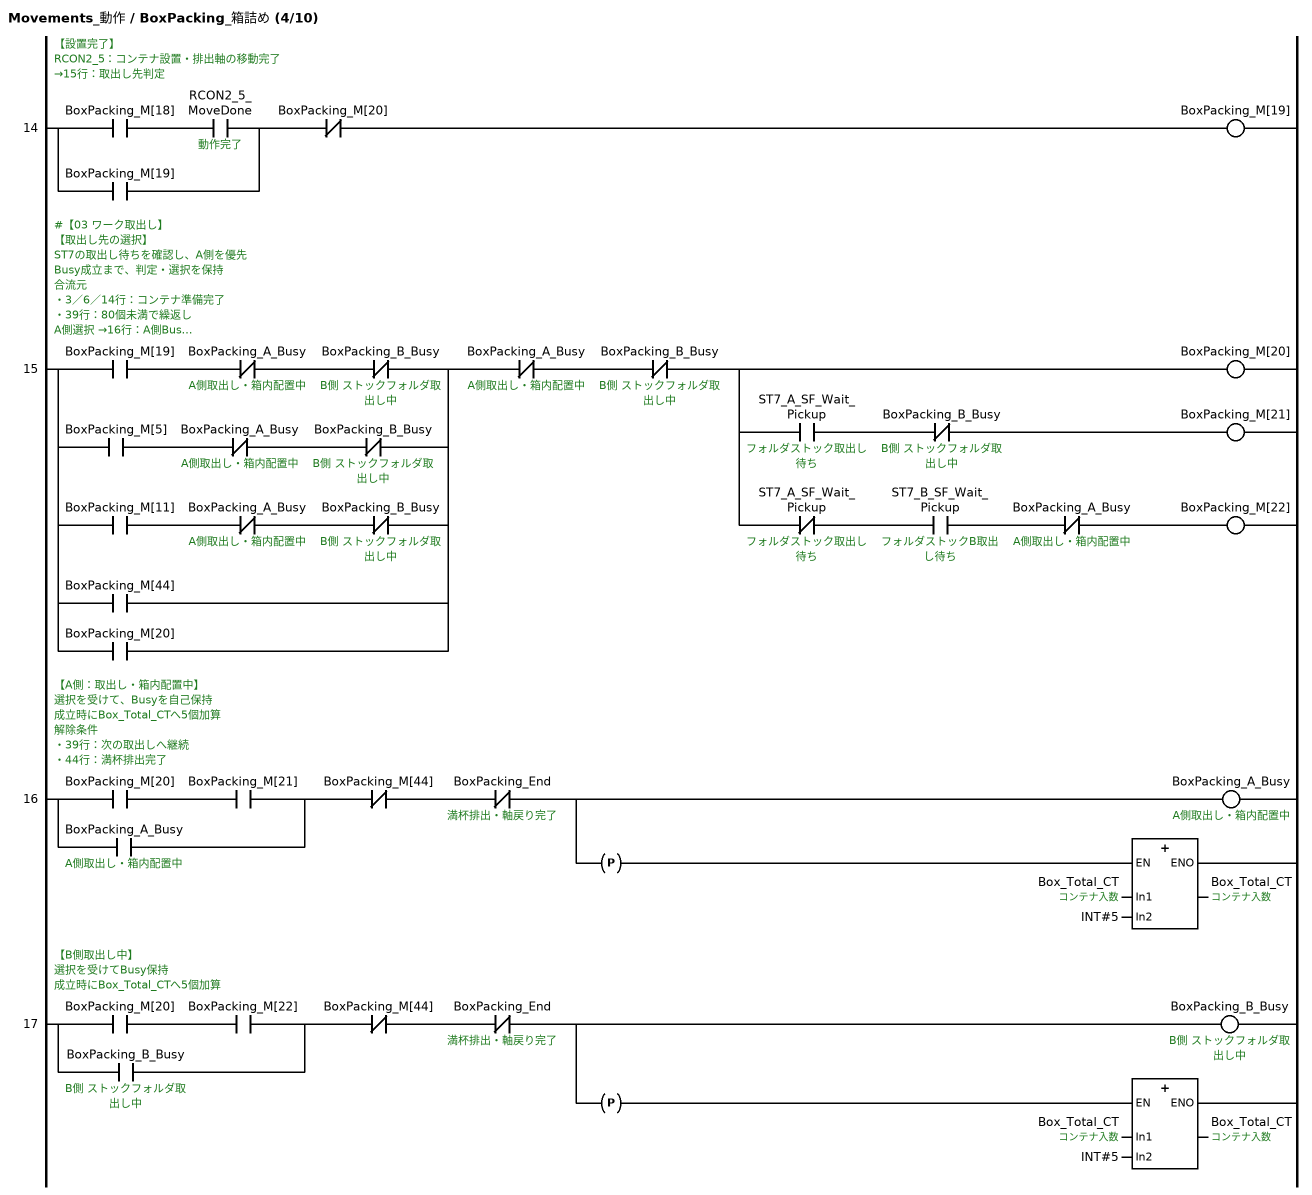
(* Rung 14: 【設置完了】 / RCON2_5：コンテナ設置・排出軸の移動完了 / →15行：取出し先判定 *)
BoxPacking_M[19] := ((BoxPacking_M[18] AND RCON2_5_MoveDone) OR BoxPacking_M[19]) AND NOT BoxPacking_M[20];
(* Rung 15: #【03 ワーク取出し】 / 【取出し先の選択】 / ST7の取出し待ちを確認し、A側を優先 / Busy成立まで、判定・選択を保持 / 合流元 / ・3／6／14行：コンテナ準備完了 / ・39行：80個未満で繰返し / A側選択 →16行：A側Busy / B側選択 →17行：B側Busy *)
_p148 := ((BoxPacking_M[19] AND NOT BoxPacking_A_Busy AND NOT BoxPacking_B_Busy) OR (BoxPacking_M[5] AND NOT BoxPacking_A_Busy AND NOT BoxPacking_B_Busy) OR (BoxPacking_M[11] AND NOT BoxPacking_A_Busy AND NOT BoxPacking_B_Busy) OR BoxPacking_M[44] OR BoxPacking_M[20]) AND NOT BoxPacking_A_Busy AND NOT BoxPacking_B_Busy;
BoxPacking_M[20] := _p148;
BoxPacking_M[21] := _p148 AND ST7_A_SF_Wait_Pickup AND NOT BoxPacking_B_Busy;
BoxPacking_M[22] := _p148 AND NOT ST7_A_SF_Wait_Pickup AND ST7_B_SF_Wait_Pickup AND NOT BoxPacking_A_Busy;
(* Rung 16: 【A側：取出し・箱内配置中】 / 選択を受けて、Busyを自己保持 / 成立時にBox_Total_CTへ5個加算 / 解除条件 / ・39行：次の取出しへ継続 / ・44行：満杯排出完了 *)
_p149 := ((BoxPacking_M[20] AND BoxPacking_M[21]) OR BoxPacking_A_Busy) AND NOT BoxPacking_M[44] AND NOT BoxPacking_End;
BoxPacking_A_Busy := _p149;
_e150(CLK := _p149);
IF _e150.Q THEN Box_Total_CT := Box_Total_CT + INT#5; END_IF;
(* Rung 17: 【B側取出し中】 / 選択を受けてBusy保持 / 成立時にBox_Total_CTへ5個加算 *)
_p151 := ((BoxPacking_M[20] AND BoxPacking_M[22]) OR BoxPacking_B_Busy) AND NOT BoxPacking_M[44] AND NOT BoxPacking_End;
BoxPacking_B_Busy := _p151;
_e152(CLK := _p151);
IF _e152.Q THEN Box_Total_CT := Box_Total_CT + INT#5; END_IF;

